(* CODESYS project Syn_Visu_3.2.0.library
   Version: 3.2.0.0
   Title: SynVisu
   Placeholder: SynVisu
   Company: Syntegon Group
   DefaultNamespace: SynVisu

Project tree, tasks and I/O mapping:
  libraries: Tc2_System, * (Beckhoff Automation GmbH)
  DUTs/
    data type E_VisuComponentType
    data type E_VisuProductState
    data type E_VisuZoneKind
    data type ST_VisuCartesian
    data type ST_VisuCartesianConfig
    data type ST_VisuCartesianState
    data type ST_VisuConveyor
    data type ST_VisuConveyorConfig
    data type ST_VisuConveyorState
    data type ST_VisuDelta
    data type ST_VisuDeltaConfig
    data type ST_VisuDeltaState
    data type ST_VisuFault
    data type ST_VisuFinger
    data type ST_VisuFingerState
    data type ST_VisuGantryMover
    data type ST_VisuLimitArea
    data type ST_VisuLoopMover
    data type ST_VisuManifest
    data type ST_VisuManifestEntry
    data type ST_VisuPlanarPose
    data type ST_VisuPose
    data type ST_VisuPosition
    data type ST_VisuProduct
    data type ST_VisuProductType
    data type ST_VisuWorkingArea
    data type ST_VisuXtsGantry
    data type ST_VisuXtsGantryConfig
    data type ST_VisuXtsGantryState
    data type ST_VisuXtsLoop
    data type ST_VisuXtsLoopConfig
    data type ST_VisuXtsLoopState
    data type ST_VisuZone
  GVLs/
    global variables VISU_GlobalConst
    global variables VISU_GlobalConst_Param
  POUs/
    function block _FB_VisuCartesian [ST]: m_ApplyConfig, m_ClearFingers, m_ClearZones, m_ComponentType, m_Configure, m_SetAxes, m_SetFault, m_SetFinger, m_SetFingerState, m_SetZone
    function block _FB_VisuComponent [ST]: m_ComponentType, m_DcTime, m_Id, m_NotifyConfigChanged, m_Register
    function block _FB_VisuConveyor [ST]: m_ApplyConfig, m_BeltPosition, m_ComponentType, m_Configure, m_FindProduct, m_GetProduct, m_LatchProduct, m_MoveProduct, m_ProductCount, m_ProductPose, m_RemoveProduct, m_RemoveProductsBeyond, m_SetBeltPosition, m_SetFault, m_SetModuloBeltPosition, m_SetProductState, m_SetProductType
    function block _FB_VisuDelta [ST]: m_ApplyConfig, m_BasePose, m_ClearFingers, m_ClearLimitArea, m_ClearZones, m_ComponentType, m_Configure, m_SetFault, m_SetFinger, m_SetFingerState, m_SetLimitArea, m_SetTcp, m_SetWorkingArea, m_SetZone
    function block _FB_VisuXtsGantry [ST]: m_ApplyConfig, m_ClearFingers, m_ClearZones, m_ComponentType, m_Configure, m_SetFault, m_SetFinger, m_SetMover, m_SetMoverCount, m_SetZone, m_SetZPosition
    function block _FB_VisuXtsLoop [ST]: m_ApplyConfig, m_ClearFingers, m_ClearZones, m_ComponentType, m_Configure, m_Perimeter, m_SetFault, m_SetFinger, m_SetMover, m_SetMoverCount, m_SetZone
    function _FC_GetVersionSynVisu [ST]
*)

// DUTs/E_VisuComponentType
{attribute 'qualified_only'}
{attribute 'strict'}
TYPE E_VisuComponentType :
(
	(* Values are part of the gateway contract: append, never renumber. *)
	NONE := 0,
	CONVEYOR := 1,
	DELTA := 2,
	XTS_GANTRY := 3,
	XTS_LOOP := 4,
	CARTESIAN := 5
) UINT;
END_TYPE

// DUTs/E_VisuProductState
{attribute 'qualified_only'}
{attribute 'strict'}
TYPE E_VisuProductState :
(
	(* Values are part of the gateway contract: append, never renumber. *)
	DETECTED := 0,
	ASSIGNED := 1,
	PICKED := 2,
	REJECTED := 3,
	PLACED := 4
) UINT;
END_TYPE

// DUTs/E_VisuZoneKind
{attribute 'qualified_only'}
{attribute 'strict'}
TYPE E_VisuZoneKind :
(
	(* Values are part of the gateway contract: append, never renumber. *)
	PICK := 1,
	PLACE := 2
) UINT;
END_TYPE

// DUTs/ST_VisuCartesian
TYPE ST_VisuCartesian :
STRUCT
	(* One visualised Cartesian robot. Register the instance's symbol path in the manifest with
	   eType := E_VisuComponentType.CARTESIAN. *)
	stConfig : ST_VisuCartesianConfig; // read at discovery and after nConfigVersion changes
	stState : ST_VisuCartesianState; // read every gateway cycle
END_STRUCT
END_TYPE

// DUTs/ST_VisuCartesianConfig
TYPE ST_VisuCartesianConfig :
STRUCT
	(* Cartesian robot: two fixed rails along local +Y, a bridge travelling in Y, a carriage on it travelling in X
	   and a vertical column (Z) ending at the gripper flange. Local frame: origin at axis X = Y = 0, Z up; the
	   flange is at (X, Y, Z). *)
	stPose : ST_VisuPose; // MCS
	fXMin : LREAL; // mm, X stroke
	fXMax : LREAL; // mm
	fYMin : LREAL; // mm, Y stroke
	fYMax : LREAL; // mm
	fZMin : LREAL; // mm, Z stroke
	fZMax : LREAL; // mm
	fRailHeight : LREAL; // mm, top of the rails above the local origin; the bridge sits on them
	nZoneCount : UINT;
	aZones : ARRAY[0..VISU_GlobalConst_Param.VISU_un_MAX_ZONES - 1] OF ST_VisuZone; // pick and place zones
	nFingerCount : UINT; // 0 = no gripper definition
	aFingers : ARRAY[0..VISU_GlobalConst_Param.VISU_un_MAX_FINGERS - 1] OF ST_VisuFinger;
END_STRUCT
END_TYPE

// DUTs/ST_VisuCartesianState
TYPE ST_VisuCartesianState :
STRUCT
	nTimestamp : ULINT; // DC time of the writing cycle, ns since 2000-01-01 (set by _FB_VisuCartesian)
	fX : LREAL; // mm, actual value: the gripper flange
	fY : LREAL; // mm, actual value
	fZ : LREAL; // mm, actual value
	bGripperActive : BOOL; // used only when no fingers are configured
	aFingerStates : ARRAY[0..VISU_GlobalConst_Param.VISU_un_MAX_FINGERS - 1] OF ST_VisuFingerState; // one per configured finger
	stFault : ST_VisuFault; // fault of the robot (set by _FB_VisuCartesian.m_SetFault)
END_STRUCT
END_TYPE

// DUTs/ST_VisuConveyor
TYPE ST_VisuConveyor :
STRUCT
	(* One visualised conveyor. Register the instance's symbol path in the manifest with
	   eType := E_VisuComponentType.CONVEYOR. *)
	stConfig : ST_VisuConveyorConfig; // read at discovery and after nConfigVersion changes
	stState : ST_VisuConveyorState; // read every gateway cycle
END_STRUCT
END_TYPE

// DUTs/ST_VisuConveyorConfig
TYPE ST_VisuConveyorConfig :
STRUCT
	stPose : ST_VisuPose; // belt start on the belt surface; local +X = conveying direction
	fLength : LREAL; // mm
	fWidth : LREAL; // mm
	nProductTypeCount : UINT;
	aProductTypes : ARRAY[0..VISU_GlobalConst_Param.VISU_un_MAX_PRODUCT_TYPES - 1] OF ST_VisuProductType;
END_STRUCT
END_TYPE

// DUTs/ST_VisuConveyorState
TYPE ST_VisuConveyorState :
STRUCT
	nTimestamp : ULINT; // DC time of the writing cycle, ns since 2000-01-01 (set by _FB_VisuConveyor)
	fBeltPosition : LREAL; // continuous belt surface position, mm, no modulo (see _FB_VisuConveyor.m_SetModuloBeltPosition)
	nProductCount : UINT; // entries [0..nProductCount-1] are evaluated
	aProducts : ARRAY[0..VISU_GlobalConst_Param.VISU_un_MAX_PRODUCTS - 1] OF ST_VisuProduct;
	stFault : ST_VisuFault; // fault of the conveyor (set by _FB_VisuConveyor.m_SetFault)
END_STRUCT
END_TYPE

// DUTs/ST_VisuDelta
TYPE ST_VisuDelta :
STRUCT
	(* One visualised Delta robot. Register the instance's symbol path in the manifest with
	   eType := E_VisuComponentType.DELTA. *)
	stConfig : ST_VisuDeltaConfig; // read at discovery and after nConfigVersion changes
	stState : ST_VisuDeltaState; // read every gateway cycle
END_STRUCT
END_TYPE

// DUTs/ST_VisuDeltaConfig
TYPE ST_VisuDeltaConfig :
STRUCT
	(* Geometry the visualisation uses to derive the arm posture from the TCP.
	   Arm 1 lies along the base's local +X; arms 2 and 3 follow counter-clockwise
	   (seen from above) at 120 deg each. *)
	stPose : ST_VisuPose; // base centre in the MCS
	fBaseRadius : LREAL; // mm, base centre to shoulder joint
	fEffectorRadius : LREAL; // mm, effector centre to lower-arm joint
	fUpperArmLength : LREAL; // mm
	fLowerArmLength : LREAL; // mm
	stWorkingArea : ST_VisuWorkingArea;
	stLimitArea : ST_VisuLimitArea; // optional box that further restricts the working area
	nZoneCount : UINT;
	aZones : ARRAY[0..VISU_GlobalConst_Param.VISU_un_MAX_ZONES - 1] OF ST_VisuZone; // pick and place zones
	nFingerCount : UINT; // 0 = no gripper definition
	aFingers : ARRAY[0..VISU_GlobalConst_Param.VISU_un_MAX_FINGERS - 1] OF ST_VisuFinger;
END_STRUCT
END_TYPE

// DUTs/ST_VisuDeltaState
TYPE ST_VisuDeltaState :
STRUCT
	nTimestamp : ULINT; // DC time of the writing cycle, ns since 2000-01-01 (set by _FB_VisuDelta.m_SetTcp)
	stActualTcp : ST_VisuPosition; // MCS, effector centre (the gripper flange); the visualisation derives the arms from it
	stSetpointTcp : ST_VisuPosition; // MCS
	aFingerStates : ARRAY[0..VISU_GlobalConst_Param.VISU_un_MAX_FINGERS - 1] OF ST_VisuFingerState; // one per configured finger
	stFault : ST_VisuFault; // fault of the robot (set by _FB_VisuDelta.m_SetFault)
END_STRUCT
END_TYPE

// DUTs/ST_VisuFault
(* Fault of a component or an XTS mover: drawn red with sMessage while bActive (contract, protocol 8). *)
TYPE ST_VisuFault :
STRUCT
	bActive : BOOL; // TRUE while the fault is active
	sMessage : STRING(80); // shown to the operator; empty shows 'Fault'
END_STRUCT
END_TYPE

// DUTs/ST_VisuFinger
TYPE ST_VisuFinger :
STRUCT
	(* One gripper finger, always drawn as a cylinder. Its frame's origin is the centre of its top face; it extends
	   along its local -Z. The grip point, where a carried product's top touches, is the centre of its bottom face. *)
	fDiameter : LREAL; // mm
	fHeight : LREAL; // mm
END_STRUCT
END_TYPE

// DUTs/ST_VisuFingerState
TYPE ST_VisuFingerState :
STRUCT
	stPose : ST_VisuPose; // MCS, absolute: pose of the finger's frame (centre of its top face)
	bActive : BOOL; // the finger grips
END_STRUCT
END_TYPE

// DUTs/ST_VisuGantryMover
TYPE ST_VisuGantryMover :
STRUCT
	nId : UDINT; // unique within the gantry, > 0; referenced by a carried product's nMoverId
	bValid : BOOL; // invalid entries are not shown
	fPosition : LREAL; // mm along the track (local +Y), actual value
	fX : LREAL; // mm, X axis on the mover, actual value
	bGripperActive : BOOL; // used only when no fingers are configured
	aFingerStates : ARRAY[0..VISU_GlobalConst_Param.VISU_un_MAX_FINGERS - 1] OF ST_VisuFingerState; // one per configured finger
	stFault : ST_VisuFault; // fault of this mover
END_STRUCT
END_TYPE

// DUTs/ST_VisuLimitArea
TYPE ST_VisuLimitArea :
STRUCT
	(* Axis-aligned box in the robot frame (relative to the base centre, turned with the robot's pose) that further
	   restricts the working area, e.g. so that neighbouring robots cannot collide. *)
	fXMin : LREAL; // mm
	fXMax : LREAL; // mm
	fYMin : LREAL; // mm
	fYMax : LREAL; // mm
	fZMin : LREAL; // mm relative to the base (below the base: negative)
	fZMax : LREAL; // mm relative to the base
	bActive : BOOL; // FALSE: no limit area, the box is not drawn
END_STRUCT
END_TYPE

// DUTs/ST_VisuLoopMover
TYPE ST_VisuLoopMover :
STRUCT
	nId : UDINT; // unique within the loop, > 0; referenced by a carried product's nMoverId
	bValid : BOOL; // invalid entries are not shown
	fPosition : LREAL; // mm along the loop from the start of the lower straight, in the conveying direction
	aFingerStates : ARRAY[0..VISU_GlobalConst_Param.VISU_un_MAX_FINGERS - 1] OF ST_VisuFingerState; // one per configured finger
	stFault : ST_VisuFault; // fault of this mover
END_STRUCT
END_TYPE

// DUTs/ST_VisuManifest
TYPE ST_VisuManifest :
STRUCT
	(* Discovery entry point. The application declares one instance at the fixed symbol
	   GVL_Visu.stManifest; the gateway starts reading there. *)
	nProtocolVersion : UINT := VISU_GlobalConst.VISU_un_PROTOCOL_VERSION;
	(* Increment after any change to the manifest or to a component's stConfig. *)
	nConfigVersion : UDINT := 1;
	nCount : UINT; // entries [0..nCount-1] are evaluated
	aEntries : ARRAY[0..VISU_GlobalConst_Param.VISU_un_MAX_MANIFEST_ENTRIES - 1] OF ST_VisuManifestEntry;
END_STRUCT
END_TYPE

// DUTs/ST_VisuManifestEntry
TYPE ST_VisuManifestEntry :
STRUCT
	nId : UDINT; // unique within the manifest, > 0; used for all cross-references
	eType : E_VisuComponentType;
	sName : STRING(80); // display name
	sPath : STRING(255); // symbol path of the ST_VisuConveyor / ST_VisuDelta instance, e.g. 'MAIN.stInfeed'
END_STRUCT
END_TYPE

// DUTs/ST_VisuPlanarPose
TYPE ST_VisuPlanarPose :
STRUCT
	(* Position plus rotation about Z in the MCS, used for TCPs and product latch poses. *)
	fX : LREAL; // mm
	fY : LREAL; // mm
	fZ : LREAL; // mm
	fRz : LREAL; // degrees
END_STRUCT
END_TYPE

// DUTs/ST_VisuPose
TYPE ST_VisuPose :
STRUCT
	(* Pose in the MCS: right-handed, Z up, X in product flow direction.
	   Rotation order R = Rz(fRz) * Ry(fRy) * Rx(fRx). *)
	fX : LREAL; // mm
	fY : LREAL; // mm
	fZ : LREAL; // mm
	fRx : LREAL; // degrees
	fRy : LREAL; // degrees
	fRz : LREAL; // degrees
END_STRUCT
END_TYPE

// DUTs/ST_VisuPosition
TYPE ST_VisuPosition :
STRUCT
	(* A point in the MCS, e.g. a Delta's TCP. *)
	fX : LREAL; // mm
	fY : LREAL; // mm
	fZ : LREAL; // mm
END_STRUCT
END_TYPE

// DUTs/ST_VisuProduct
TYPE ST_VisuProduct :
STRUCT
	nId : UDINT;
	bValid : BOOL; // invalid entries are not shown
	stLatchPose : ST_VisuPlanarPose; // MCS, bottom centre of the product at latch time
	fLatchBeltPosition : LREAL; // conveyor fBeltPosition at latch time, mm
	eState : E_VisuProductState;
	nRobotId : UDINT; // manifest id of the assigned robot, 0 = none
	nMoverId : UDINT; // mover of an XTS gantry or loop carrying the product, 0 = none
	nFingerId : UDINT; // gripper finger (1-based) the product hangs from while picked, 0 = the gripper flange
	nProductType : UDINT; // id in the conveyor's aProductTypes
END_STRUCT
END_TYPE

// DUTs/ST_VisuProductType
TYPE ST_VisuProductType :
STRUCT
	nId : UDINT;
	fLength : LREAL; // mm, along the conveying direction
	fWidth : LREAL; // mm
	fHeight : LREAL; // mm
END_STRUCT
END_TYPE

// DUTs/ST_VisuWorkingArea
TYPE ST_VisuWorkingArea :
STRUCT
	(* Limit shape the PLC enforces: vertical cylinder in the robot frame, optional cone below. *)
	fRadius : LREAL; // mm
	fZMin : LREAL; // mm relative to the base (below the base: negative)
	fZMax : LREAL; // mm relative to the base
	fConeHeight : LREAL; // mm below fZMin; 0 = no cone
	fConeBottomRadius : LREAL; // mm
END_STRUCT
END_TYPE

// DUTs/ST_VisuXtsGantry
TYPE ST_VisuXtsGantry :
STRUCT
	(* One visualised XTS gantry (e.g. IDH). Register the instance's symbol path in the manifest with
	   eType := E_VisuComponentType.XTS_GANTRY. *)
	stConfig : ST_VisuXtsGantryConfig; // read at discovery and after nConfigVersion changes
	stState : ST_VisuXtsGantryState; // read every gateway cycle
END_STRUCT
END_TYPE

// DUTs/ST_VisuXtsGantryConfig
TYPE ST_VisuXtsGantryConfig :
STRUCT
	(* Straight XTS track of equal modules, carried by a common Z axis; every mover carries an X axis with a
	   gripper flange at its end. Local frame: origin at the track start on top of the movers with Z = 0; the track runs
	   along local +Y, the X axes along local +X, the Z axis along local +Z (up). *)
	stPose : ST_VisuPose; // MCS
	nModuleCount : UINT; // track modules in a row
	fModuleLength : LREAL; // mm, length of one module
	fXMin : LREAL; // mm, X stroke
	fXMax : LREAL; // mm
	fZMin : LREAL; // mm, Z stroke
	fZMax : LREAL; // mm
	fToolOffsetX : LREAL; // mm, gripper flange ahead of the X axis zero along local +X
	fToolOffsetZ : LREAL; // mm, gripper flange relative to the mover top (below: negative)
	fMoverLength : LREAL; // mm, along the track
	fMoverWidth : LREAL; // mm
	nZoneCount : UINT;
	aZones : ARRAY[0..VISU_GlobalConst_Param.VISU_un_MAX_ZONES - 1] OF ST_VisuZone; // pick and place zones
	nFingerCount : UINT; // fingers of every mover's gripper, 0 = no gripper definition
	aFingers : ARRAY[0..VISU_GlobalConst_Param.VISU_un_MAX_FINGERS - 1] OF ST_VisuFinger;
END_STRUCT
END_TYPE

// DUTs/ST_VisuXtsGantryState
TYPE ST_VisuXtsGantryState :
STRUCT
	nTimestamp : ULINT; // DC time of the writing cycle, ns since 2000-01-01 (set by _FB_VisuXtsGantry)
	fZ : LREAL; // mm, common Z axis, actual value
	nMoverCount : UINT; // entries [0..nMoverCount-1] are evaluated
	aMovers : ARRAY[0..VISU_GlobalConst_Param.VISU_un_MAX_MOVERS - 1] OF ST_VisuGantryMover;
	stFault : ST_VisuFault; // fault of the whole gantry (set by _FB_VisuXtsGantry.m_SetFault)
END_STRUCT
END_TYPE

// DUTs/ST_VisuXtsLoop
TYPE ST_VisuXtsLoop :
STRUCT
	(* One visualised XTS loop (e.g. Fxx). Register the instance's symbol path in the manifest with
	   eType := E_VisuComponentType.XTS_LOOP. *)
	stConfig : ST_VisuXtsLoopConfig; // read at discovery and after nConfigVersion changes
	stState : ST_VisuXtsLoopState; // read every gateway cycle
END_STRUCT
END_TYPE

// DUTs/ST_VisuXtsLoopConfig
TYPE ST_VisuXtsLoopConfig :
STRUCT
	(* Closed XTS loop: two straights joined by two 180 deg curves (drawn as semicircles), standing in the local X-Z
	   plane. Local frame: origin at the start of the lower straight, which runs along local +X in the conveying
	   direction; the upper straight lies at +2 * fCurveRadius in Z. *)
	stPose : ST_VisuPose; // MCS
	fStraightLength : LREAL; // mm
	fCurveRadius : LREAL; // mm
	fToolOffset : LREAL; // mm, gripper flange (tool point) of a mover outwards from the track
	fMoverLength : LREAL; // mm, along the track
	fMoverWidth : LREAL; // mm
	nZoneCount : UINT;
	aZones : ARRAY[0..VISU_GlobalConst_Param.VISU_un_MAX_ZONES - 1] OF ST_VisuZone; // pick and place zones
	nFingerCount : UINT; // fingers of every mover's gripper, 0 = no gripper definition
	aFingers : ARRAY[0..VISU_GlobalConst_Param.VISU_un_MAX_FINGERS - 1] OF ST_VisuFinger;
END_STRUCT
END_TYPE

// DUTs/ST_VisuXtsLoopState
TYPE ST_VisuXtsLoopState :
STRUCT
	nTimestamp : ULINT; // DC time of the writing cycle, ns since 2000-01-01 (set by _FB_VisuXtsLoop)
	nMoverCount : UINT; // entries [0..nMoverCount-1] are evaluated
	aMovers : ARRAY[0..VISU_GlobalConst_Param.VISU_un_MAX_MOVERS - 1] OF ST_VisuLoopMover;
	stFault : ST_VisuFault; // fault of the whole loop (set by _FB_VisuXtsLoop.m_SetFault)
END_STRUCT
END_TYPE

// DUTs/ST_VisuZone
TYPE ST_VisuZone :
STRUCT
	nConveyorId : UDINT; // manifest id of the conveyor
	fStart : LREAL; // mm along the conveyor's local X (belt coordinates, not MCS)
	fEnd : LREAL; // mm along the conveyor's local X
	eKind : E_VisuZoneKind;
	(* mm before fEnd, against the conveying direction: the robot may allocate products in the zone only up to
	   fEnd - fAllocationOffset, so it does not move out of the zone while approaching. 0 = no allocation limit. *)
	fAllocationOffset : LREAL;
END_STRUCT
END_TYPE

// GVLs/VISU_GlobalConst
(****************************************************************************************************<br>
© Syntegon Group.<br>
All rights reserved, also regarding any disposal, exploitation, reproduction, editing, distribution,<br>
as well as in the event of applications for industrial property rights.<br>
*****************************************************************************************************<br>
DESCRIPTION:<br>
Global constants of the Syn_Visu library.<br>
****************************************************************************************************)
{attribute 'qualified_only'}
VAR_GLOBAL CONSTANT
	(* Version of the PLC <-> gateway contract. The gateway refuses to read a PLC whose manifest
	   reports a different value. Bump together with PROTOCOL_VERSION in the gateway.
	   2: the Delta reports only its TCP; the visualisation derives the arm posture.
	   3: work area renamed to working area, windows to zones.
	   4: XTS gantry and XTS loop, product nMoverId, fEncoder renamed to fBeltPosition.
	   5: Cartesian robot.
	   6: Delta limit area, zone allocation offset.
	   7: gripper fingers; tool rotations (Delta rz, IDH C, Cartesian C/A and tool length) removed.
	   8: faults of components and XTS movers (stFault). *)
	VISU_un_PROTOCOL_VERSION			: UINT := 8;
	VISU_lr_DEG_TO_RAD					: LREAL := 0.017453292519943295;	// [rad/deg] pi / 180
END_VAR

// GVLs/VISU_GlobalConst_Param
(****************************************************************************************************<br>
© Syntegon Group.<br>
All rights reserved, also regarding any disposal, exploitation, reproduction, editing, distribution,<br>
as well as in the event of applications for industrial property rights.<br>
*****************************************************************************************************<br>
DESCRIPTION:<br>
Library parameters of Syn_Visu: array sizes of the interface structures.<br>
****************************************************************************************************)
{attribute 'qualified_only'}
VAR_GLOBAL CONSTANT
	VISU_un_MAX_MANIFEST_ENTRIES		: UINT := 32;	// [-] components in the manifest
	VISU_un_MAX_PRODUCTS				: UINT := 128;	// [-] products per conveyor
	VISU_un_MAX_PRODUCT_TYPES			: UINT := 8;	// [-] product types per conveyor
	VISU_un_MAX_ZONES					: UINT := 8;	// [-] zones per robot
	VISU_un_MAX_MOVERS					: UINT := 40;	// [-] movers per XTS gantry or loop
	VISU_un_MAX_FINGERS					: UINT := 8;	// [-] fingers per gripper
END_VAR

// POUs/_FB_VisuCartesian
(****************************************************************************************************<br>
© Syntegon Group.<br>
All rights reserved, also regarding any disposal, exploitation, reproduction, editing, distribution,<br>
as well as in the event of applications for industrial property rights.<br>
*****************************************************************************************************<br>
DESCRIPTION:<br>
One visualised Cartesian robot: linear X, Y, Z axes ending at a gripper flange. Typical cycle:<br>
  fb_Cartesian.m_Register(vio_Manifest := GVL_Visu.stManifest, vi_udn_Id := 40, vi_str_Name := 'Cartesian',<br>
      vi_str_Path := 'MAIN.fb_Cartesian.vo_Visu');<br>
  fb_Cartesian.m_Configure(vi_Pose := RobotPose, vi_lr_XMin := 0, vi_lr_XMax := 1200, vi_lr_YMin := 0,<br>
      vi_lr_YMax := 1000, vi_lr_ZMin := -600, vi_lr_ZMax := 0, vi_lr_RailHeight := 1200);<br>
  fb_Cartesian.m_SetFinger(vi_un_Finger := 1, vi_lr_Diameter := 40, vi_lr_Height := 40);<br>
  fb_Cartesian.m_SetZone(vi_udn_ConveyorId := 7, vi_e_Kind := E_VisuZoneKind.PICK, vi_lr_Start := 1000, vi_lr_End := 2000);<br>
  fb_Cartesian.m_SetAxes(vi_lr_X := ..., vi_lr_Y := ..., vi_lr_Z := ...);<br>
  fb_Cartesian.m_SetFingerState(vi_un_Finger := 1, vi_Pose := CupPose, vi_b_Active := b_Vacuum);<br>
Only actual values are reported; tool rotations (e.g. C and A) show only through the finger poses, absolute in<br>
the MCS. The config methods may be called every cycle; the config version only changes when a value does.<br>
*****************************************************************************************************<br>
OUTPUT VALUES:<br>
vo_Visu is the contract structure the gateway reads at the path given to m_Register. Do not write it.<br>
*****************************************************************************************************<br>
VERSION         ¦ DATE       ¦ NAME      ¦ CHANGE<br>
Syn_Visu 3.0.0  ¦ 2026-10-31 ¦ J.Willner ¦ Naming and layout after the TCAT programming guideline<br>
****************************************************************************************************)
FUNCTION_BLOCK _FB_VisuCartesian EXTENDS _FB_VisuComponent
VAR_OUTPUT
	vo_Visu								: ST_VisuCartesian;	// contract structure read by the gateway
END_VAR

(****************************************************************************************************<br>
© Syntegon Group.<br>
All rights reserved, also regarding any disposal, exploitation, reproduction, editing, distribution,<br>
as well as in the event of applications for industrial property rights.<br>
*****************************************************************************************************<br>
DESCRIPTION:<br>
Takes over vio_New and increments the config version if it differs from the current config. TRUE if changed.<br>
****************************************************************************************************)
METHOD PRIVATE m_ApplyConfig : BOOL
VAR_IN_OUT
	vio_New								: ST_VisuCartesianConfig;
END_VAR
m_ApplyConfig := Tc2_System.MEMCMP(ADR(vio_New), ADR(vo_Visu.stConfig), SIZEOF(vio_New)) <> 0;
IF m_ApplyConfig THEN
	vo_Visu.stConfig := vio_New;
	m_NotifyConfigChanged();
END_IF
END_METHOD

(****************************************************************************************************<br>
© Syntegon Group.<br>
All rights reserved, also regarding any disposal, exploitation, reproduction, editing, distribution,<br>
as well as in the event of applications for industrial property rights.<br>
*****************************************************************************************************<br>
DESCRIPTION:<br>
Removes the gripper definition. TRUE if there was one.<br>
****************************************************************************************************)
METHOD m_ClearFingers : BOOL
VAR
	TempNew								: ST_VisuCartesianConfig;
	TempEmpty							: ST_VisuFinger;
	un_TempIndex						: UINT;
END_VAR
TempNew := vo_Visu.stConfig;
FOR un_TempIndex := 0 TO VISU_GlobalConst_Param.VISU_un_MAX_FINGERS - 1 DO
	TempNew.aFingers[un_TempIndex] := TempEmpty;
END_FOR
TempNew.nFingerCount := 0;
m_ClearFingers := m_ApplyConfig(TempNew);
END_METHOD

(****************************************************************************************************<br>
© Syntegon Group.<br>
All rights reserved, also regarding any disposal, exploitation, reproduction, editing, distribution,<br>
as well as in the event of applications for industrial property rights.<br>
*****************************************************************************************************<br>
DESCRIPTION:<br>
Removes all pick and place zones. TRUE if there were any.<br>
****************************************************************************************************)
METHOD m_ClearZones : BOOL
VAR
	TempNew								: ST_VisuCartesianConfig;
	TempEmpty							: ST_VisuZone;
	un_TempIndex						: UINT;
END_VAR
TempNew := vo_Visu.stConfig;
FOR un_TempIndex := 0 TO VISU_GlobalConst_Param.VISU_un_MAX_ZONES - 1 DO
	TempNew.aZones[un_TempIndex] := TempEmpty;
END_FOR
TempNew.nZoneCount := 0;
m_ClearZones := m_ApplyConfig(TempNew);
END_METHOD

(****************************************************************************************************<br>
© Syntegon Group.<br>
All rights reserved, also regarding any disposal, exploitation, reproduction, editing, distribution,<br>
as well as in the event of applications for industrial property rights.<br>
*****************************************************************************************************<br>
DESCRIPTION:<br>
Manifest type: Cartesian robot.<br>
****************************************************************************************************)
METHOD PROTECTED m_ComponentType : E_VisuComponentType
m_ComponentType := E_VisuComponentType.CARTESIAN;
END_METHOD

(****************************************************************************************************<br>
© Syntegon Group.<br>
All rights reserved, also regarding any disposal, exploitation, reproduction, editing, distribution,<br>
as well as in the event of applications for industrial property rights.<br>
*****************************************************************************************************<br>
DESCRIPTION:<br>
Sets pose, strokes and rail height. TRUE if anything changed.<br>
****************************************************************************************************)
METHOD m_Configure : BOOL
VAR_INPUT
	vi_Pose								: ST_VisuPose;	// MCS, axis origin X = Y = 0 with Z up
	vi_lr_XMin							: LREAL;	// [mm]
	vi_lr_XMax							: LREAL;	// [mm]
	vi_lr_YMin							: LREAL;	// [mm]
	vi_lr_YMax							: LREAL;	// [mm]
	vi_lr_ZMin							: LREAL;	// [mm]
	vi_lr_ZMax							: LREAL;	// [mm]
	vi_lr_RailHeight					: LREAL;	// [mm] top of the rails above the local origin
END_VAR
VAR
	TempNew								: ST_VisuCartesianConfig;
END_VAR
TempNew := vo_Visu.stConfig;
TempNew.stPose := vi_Pose;
TempNew.fXMin := vi_lr_XMin;
TempNew.fXMax := vi_lr_XMax;
TempNew.fYMin := vi_lr_YMin;
TempNew.fYMax := vi_lr_YMax;
TempNew.fZMin := vi_lr_ZMin;
TempNew.fZMax := vi_lr_ZMax;
TempNew.fRailHeight := vi_lr_RailHeight;
m_Configure := m_ApplyConfig(TempNew);
END_METHOD

(****************************************************************************************************<br>
© Syntegon Group.<br>
All rights reserved, also regarding any disposal, exploitation, reproduction, editing, distribution,<br>
as well as in the event of applications for industrial property rights.<br>
*****************************************************************************************************<br>
DESCRIPTION:<br>
Reports the axes' actual values and the gripper. Call once per cycle; it also stamps the state with the<br>
cycle's DC time.<br>
****************************************************************************************************)
METHOD m_SetAxes : BOOL
VAR_INPUT
	vi_lr_X								: LREAL;	// [mm]
	vi_lr_Y								: LREAL;	// [mm]
	vi_lr_Z								: LREAL;	// [mm]
	vi_b_GripperActive					: BOOL := FALSE;	// used only when no fingers are configured
END_VAR
vo_Visu.stState.fX := vi_lr_X;
vo_Visu.stState.fY := vi_lr_Y;
vo_Visu.stState.fZ := vi_lr_Z;
vo_Visu.stState.bGripperActive := vi_b_GripperActive;
vo_Visu.stState.nTimestamp := m_DcTime();
m_SetAxes := TRUE;
END_METHOD

(****************************************************************************************************<br>
© Syntegon Group.<br>
All rights reserved, also regarding any disposal, exploitation, reproduction, editing, distribution,<br>
as well as in the event of applications for industrial property rights.<br>
*****************************************************************************************************<br>
DESCRIPTION:<br>
Sets or clears the fault of the robot: drawn red with the message while active. The fault stays until it<br>
is cleared with m_SetFault(vi_b_Active := FALSE, vi_str_Message := ''). TRUE.<br>
****************************************************************************************************)
METHOD m_SetFault : BOOL
VAR_INPUT
	vi_b_Active							: BOOL;	// TRUE: fault active
	vi_str_Message						: STRING(80);	// shown to the operator; empty shows 'Fault'
END_VAR
vo_Visu.stState.stFault.bActive := vi_b_Active;
vo_Visu.stState.stFault.sMessage := vi_str_Message;
m_SetFault := TRUE;
END_METHOD

(****************************************************************************************************<br>
© Syntegon Group.<br>
All rights reserved, also regarding any disposal, exploitation, reproduction, editing, distribution,<br>
as well as in the event of applications for industrial property rights.<br>
*****************************************************************************************************<br>
DESCRIPTION:<br>
Defines gripper finger vi_un_Finger (1-based): a cylinder hanging from the finger's pose along its local -Z.<br>
The finger count grows to vi_un_Finger.<br>
*****************************************************************************************************<br>
OUTPUT VALUES:<br>
FALSE outside 1..VISU_GlobalConst_Param.VISU_un_MAX_FINGERS.<br>
****************************************************************************************************)
METHOD m_SetFinger : BOOL
VAR_INPUT
	vi_un_Finger						: UINT;	// [-] 1-based, as a product's nFingerId
	vi_lr_Diameter						: LREAL;	// [mm]
	vi_lr_Height						: LREAL;	// [mm] along the finger's local -Z
END_VAR
VAR
	TempNew								: ST_VisuCartesianConfig;
END_VAR
m_SetFinger := FALSE;
IF vi_un_Finger = 0 OR vi_un_Finger > VISU_GlobalConst_Param.VISU_un_MAX_FINGERS THEN
	RETURN;
END_IF
TempNew := vo_Visu.stConfig;
TempNew.aFingers[vi_un_Finger - 1].fDiameter := vi_lr_Diameter;
TempNew.aFingers[vi_un_Finger - 1].fHeight := vi_lr_Height;
TempNew.nFingerCount := MAX(TempNew.nFingerCount, vi_un_Finger);
m_ApplyConfig(TempNew);
m_SetFinger := TRUE;
END_METHOD

(****************************************************************************************************<br>
© Syntegon Group.<br>
All rights reserved, also regarding any disposal, exploitation, reproduction, editing, distribution,<br>
as well as in the event of applications for industrial property rights.<br>
*****************************************************************************************************<br>
DESCRIPTION:<br>
Reports finger vi_un_Finger (1-based): the pose of its frame (centre of its top face), absolute in the MCS,<br>
and whether it grips. Call once per cycle per configured finger.<br>
*****************************************************************************************************<br>
OUTPUT VALUES:<br>
FALSE outside 1..VISU_GlobalConst_Param.VISU_un_MAX_FINGERS.<br>
****************************************************************************************************)
METHOD m_SetFingerState : BOOL
VAR_INPUT
	vi_un_Finger						: UINT;	// [-] 1-based
	vi_Pose								: ST_VisuPose;	// MCS
	vi_b_Active							: BOOL;	// TRUE while the finger grips
END_VAR
m_SetFingerState := vi_un_Finger > 0 AND vi_un_Finger <= VISU_GlobalConst_Param.VISU_un_MAX_FINGERS;
IF m_SetFingerState THEN
	vo_Visu.stState.aFingerStates[vi_un_Finger - 1].stPose := vi_Pose;
	vo_Visu.stState.aFingerStates[vi_un_Finger - 1].bActive := vi_b_Active;
END_IF
END_METHOD

(****************************************************************************************************<br>
© Syntegon Group.<br>
All rights reserved, also regarding any disposal, exploitation, reproduction, editing, distribution,<br>
as well as in the event of applications for industrial property rights.<br>
*****************************************************************************************************<br>
DESCRIPTION:<br>
Adds a pick or place zone, or updates the one for the same conveyor and kind.<br>
*****************************************************************************************************<br>
OUTPUT VALUES:<br>
FALSE for vi_udn_ConveyorId = 0 or a full list.<br>
****************************************************************************************************)
METHOD m_SetZone : BOOL
VAR_INPUT
	vi_udn_ConveyorId					: UDINT;	// [-] manifest id of the conveyor
	vi_e_Kind							: E_VisuZoneKind;
	vi_lr_Start							: LREAL;	// [mm] along the conveyor from its start (belt coordinates, not MCS)
	vi_lr_End							: LREAL;	// [mm] along the conveyor from its start
	vi_lr_AllocationOffset				: LREAL := 0;	// [mm] before vi_lr_End up to which products may be allocated; 0 = no limit
END_VAR
VAR
	TempNew								: ST_VisuCartesianConfig;
	un_TempIndex						: UINT;
END_VAR
m_SetZone := FALSE;
IF vi_udn_ConveyorId = 0 THEN
	RETURN;
END_IF
TempNew := vo_Visu.stConfig;
un_TempIndex := 0;
(* ST evaluates both operands of AND: test the index before reading the array. *)
WHILE un_TempIndex < TempNew.nZoneCount DO
	IF TempNew.aZones[un_TempIndex].nConveyorId = vi_udn_ConveyorId AND TempNew.aZones[un_TempIndex].eKind = vi_e_Kind THEN
		EXIT;
	END_IF
	un_TempIndex := un_TempIndex + 1;
END_WHILE
IF un_TempIndex >= VISU_GlobalConst_Param.VISU_un_MAX_ZONES THEN
	RETURN;
END_IF
IF un_TempIndex = TempNew.nZoneCount THEN
	TempNew.nZoneCount := TempNew.nZoneCount + 1;
END_IF
TempNew.aZones[un_TempIndex].nConveyorId := vi_udn_ConveyorId;
TempNew.aZones[un_TempIndex].eKind := vi_e_Kind;
TempNew.aZones[un_TempIndex].fStart := vi_lr_Start;
TempNew.aZones[un_TempIndex].fEnd := vi_lr_End;
TempNew.aZones[un_TempIndex].fAllocationOffset := vi_lr_AllocationOffset;
m_ApplyConfig(TempNew);
m_SetZone := TRUE;
END_METHOD

END_FUNCTION_BLOCK

// POUs/_FB_VisuComponent
(****************************************************************************************************<br>
© Syntegon Group.<br>
All rights reserved, also regarding any disposal, exploitation, reproduction, editing, distribution,<br>
as well as in the event of applications for industrial property rights.<br>
*****************************************************************************************************<br>
DESCRIPTION:<br>
Base of every visualised component (_FB_VisuConveyor, _FB_VisuDelta, ...). Handles the manifest entry,<br>
the config version and the DC timestamps. Not used directly.<br>
*****************************************************************************************************<br>
VERSION         ¦ DATE       ¦ NAME      ¦ CHANGE<br>
Syn_Visu 3.0.0  ¦ 2026-10-31 ¦ J.Willner ¦ Naming and layout after the TCAT programming guideline<br>
****************************************************************************************************)
FUNCTION_BLOCK ABSTRACT _FB_VisuComponent
VAR
	RefManifest							: REFERENCE TO ST_VisuManifest;	// set by m_Register
	udn_ComponentId						: UDINT;	// [-] manifest id, 0 = not registered
END_VAR

(****************************************************************************************************<br>
© Syntegon Group.<br>
All rights reserved, also regarding any disposal, exploitation, reproduction, editing, distribution,<br>
as well as in the event of applications for industrial property rights.<br>
*****************************************************************************************************<br>
DESCRIPTION:<br>
Manifest type of the component. Overridden by every derived FB.<br>
****************************************************************************************************)
METHOD PROTECTED m_ComponentType : E_VisuComponentType
m_ComponentType := E_VisuComponentType.NONE;
END_METHOD

(****************************************************************************************************<br>
© Syntegon Group.<br>
All rights reserved, also regarding any disposal, exploitation, reproduction, editing, distribution,<br>
as well as in the event of applications for industrial property rights.<br>
*****************************************************************************************************<br>
DESCRIPTION:<br>
Distributed-clock time of the calling task's current cycle in ns since 2000-01-01; 0 if unknown.<br>
****************************************************************************************************)
METHOD PROTECTED m_DcTime : ULINT
VAR
	dn_TempTaskIndex					: DINT;
END_VAR
dn_TempTaskIndex := Tc2_System.GETCURTASKINDEXEX();
IF dn_TempTaskIndex > 0 THEN
	m_DcTime := LINT_TO_ULINT(TwinCAT_SystemInfoVarList._TaskInfo[dn_TempTaskIndex].DcTaskTime);
ELSE
	m_DcTime := 0;
END_IF
END_METHOD

(****************************************************************************************************<br>
© Syntegon Group.<br>
All rights reserved, also regarding any disposal, exploitation, reproduction, editing, distribution,<br>
as well as in the event of applications for industrial property rights.<br>
*****************************************************************************************************<br>
DESCRIPTION:<br>
Manifest id given to m_Register; 0 while not registered.<br>
****************************************************************************************************)
METHOD m_Id : UDINT
m_Id := udn_ComponentId;
END_METHOD

(****************************************************************************************************<br>
© Syntegon Group.<br>
All rights reserved, also regarding any disposal, exploitation, reproduction, editing, distribution,<br>
as well as in the event of applications for industrial property rights.<br>
*****************************************************************************************************<br>
DESCRIPTION:<br>
Increments the manifest's nConfigVersion so the gateway re-reads the config. No effect before m_Register.<br>
****************************************************************************************************)
METHOD PROTECTED m_NotifyConfigChanged : BOOL
m_NotifyConfigChanged := __ISVALIDREF(RefManifest);
IF m_NotifyConfigChanged THEN
	RefManifest.nConfigVersion := RefManifest.nConfigVersion + 1;
END_IF
END_METHOD

(****************************************************************************************************<br>
© Syntegon Group.<br>
All rights reserved, also regarding any disposal, exploitation, reproduction, editing, distribution,<br>
as well as in the event of applications for industrial property rights.<br>
*****************************************************************************************************<br>
DESCRIPTION:<br>
Adds this component to the manifest; increments nConfigVersion when the entry is new.<br>
Idempotent: call it every cycle, which also keeps the manifest reference valid after an online change.<br>
*****************************************************************************************************<br>
OUTPUT VALUES:<br>
FALSE for vi_udn_Id = 0, an id already used by a different entry, or a full manifest.<br>
****************************************************************************************************)
METHOD m_Register : BOOL
VAR_IN_OUT
	vio_Manifest						: ST_VisuManifest;	// GVL_Visu.stManifest of the application
END_VAR
VAR_INPUT
	vi_udn_Id							: UDINT;	// [-] unique, > 0
	vi_str_Name							: STRING(80);	// display name
	vi_str_Path							: STRING(255);	// symbol path of this instance's vo_Visu, e.g. 'MAIN.fb_Infeed.vo_Visu'
END_VAR
VAR
	e_TempType							: E_VisuComponentType;
	un_TempIndex						: UINT;
END_VAR
m_Register := FALSE;
RefManifest REF= vio_Manifest;
(* Always report the contract version of the library actually running, also after an online change. *)
vio_Manifest.nProtocolVersion := VISU_GlobalConst.VISU_un_PROTOCOL_VERSION;
e_TempType := m_ComponentType();
IF vi_udn_Id = 0 OR e_TempType = E_VisuComponentType.NONE THEN
	RETURN;
END_IF

(* An existing entry with the same id must match exactly. *)
un_TempIndex := 0;
WHILE un_TempIndex < vio_Manifest.nCount AND un_TempIndex < VISU_GlobalConst_Param.VISU_un_MAX_MANIFEST_ENTRIES DO
	IF vio_Manifest.aEntries[un_TempIndex].nId = vi_udn_Id THEN
		m_Register := vio_Manifest.aEntries[un_TempIndex].eType = e_TempType
					AND vio_Manifest.aEntries[un_TempIndex].sName = vi_str_Name
					AND vio_Manifest.aEntries[un_TempIndex].sPath = vi_str_Path;
		IF m_Register THEN
			udn_ComponentId := vi_udn_Id;
		END_IF
		RETURN;
	END_IF
	un_TempIndex := un_TempIndex + 1;
END_WHILE

(* New entry. *)
IF vio_Manifest.nCount >= VISU_GlobalConst_Param.VISU_un_MAX_MANIFEST_ENTRIES THEN
	RETURN;
END_IF
vio_Manifest.aEntries[vio_Manifest.nCount].nId := vi_udn_Id;
vio_Manifest.aEntries[vio_Manifest.nCount].eType := e_TempType;
vio_Manifest.aEntries[vio_Manifest.nCount].sName := vi_str_Name;
vio_Manifest.aEntries[vio_Manifest.nCount].sPath := vi_str_Path;
vio_Manifest.nCount := vio_Manifest.nCount + 1;
vio_Manifest.nConfigVersion := vio_Manifest.nConfigVersion + 1;
udn_ComponentId := vi_udn_Id;
m_Register := TRUE;
END_METHOD

END_FUNCTION_BLOCK

// POUs/_FB_VisuConveyor
(****************************************************************************************************<br>
© Syntegon Group.<br>
All rights reserved, also regarding any disposal, exploitation, reproduction, editing, distribution,<br>
as well as in the event of applications for industrial property rights.<br>
*****************************************************************************************************<br>
DESCRIPTION:<br>
One visualised conveyor. Typical cycle:<br>
  fb_Infeed.m_Register(vio_Manifest := GVL_Visu.stManifest, vi_udn_Id := 1, vi_str_Name := 'Infeed',<br>
      vi_str_Path := 'MAIN.fb_Infeed.vo_Visu');<br>
  fb_Infeed.m_Configure(vi_Pose := BeltPose, vi_lr_Length := 5000, vi_lr_Width := 400);<br>
  fb_Infeed.m_SetProductType(vi_udn_Id := 1, vi_lr_Length := 120, vi_lr_Width := 80, vi_lr_Height := 40);<br>
  fb_Infeed.m_SetBeltPosition(lr_AxisPosition);  // or m_SetModuloBeltPosition for a modulo axis<br>
  IF b_Latched THEN fb_Infeed.m_LatchProduct(vi_udn_Id := udn_NextId, vi_LatchPose := LatchPose, vi_udn_ProductType := 1); END_IF<br>
m_Configure and m_SetProductType may be called every cycle; the config version only changes when a value does.<br>
*****************************************************************************************************<br>
OUTPUT VALUES:<br>
vo_Visu is the contract structure the gateway reads at the path given to m_Register. Do not write it.<br>
*****************************************************************************************************<br>
VERSION         ¦ DATE       ¦ NAME      ¦ CHANGE<br>
Syn_Visu 3.0.0  ¦ 2026-10-31 ¦ J.Willner ¦ Naming and layout after the TCAT programming guideline<br>
****************************************************************************************************)
FUNCTION_BLOCK _FB_VisuConveyor EXTENDS _FB_VisuComponent
VAR_OUTPUT
	vo_Visu								: ST_VisuConveyor;	// contract structure read by the gateway
END_VAR
VAR
	lr_LastModuloPosition				: LREAL;	// [mm] modulo position of the previous cycle
	b_ModuloInitialised					: BOOL;
END_VAR

(****************************************************************************************************<br>
© Syntegon Group.<br>
All rights reserved, also regarding any disposal, exploitation, reproduction, editing, distribution,<br>
as well as in the event of applications for industrial property rights.<br>
*****************************************************************************************************<br>
DESCRIPTION:<br>
Takes over vio_New and increments the config version if it differs from the current config. TRUE if changed.<br>
****************************************************************************************************)
METHOD PRIVATE m_ApplyConfig : BOOL
VAR_IN_OUT
	vio_New								: ST_VisuConveyorConfig;
END_VAR
m_ApplyConfig := Tc2_System.MEMCMP(ADR(vio_New), ADR(vo_Visu.stConfig), SIZEOF(vio_New)) <> 0;
IF m_ApplyConfig THEN
	vo_Visu.stConfig := vio_New;
	m_NotifyConfigChanged();
END_IF
END_METHOD

(****************************************************************************************************<br>
© Syntegon Group.<br>
All rights reserved, also regarding any disposal, exploitation, reproduction, editing, distribution,<br>
as well as in the event of applications for industrial property rights.<br>
*****************************************************************************************************<br>
DESCRIPTION:<br>
Belt position last set, [mm].<br>
****************************************************************************************************)
METHOD m_BeltPosition : LREAL
m_BeltPosition := vo_Visu.stState.fBeltPosition;
END_METHOD

(****************************************************************************************************<br>
© Syntegon Group.<br>
All rights reserved, also regarding any disposal, exploitation, reproduction, editing, distribution,<br>
as well as in the event of applications for industrial property rights.<br>
*****************************************************************************************************<br>
DESCRIPTION:<br>
Manifest type: conveyor.<br>
****************************************************************************************************)
METHOD PROTECTED m_ComponentType : E_VisuComponentType
m_ComponentType := E_VisuComponentType.CONVEYOR;
END_METHOD

(****************************************************************************************************<br>
© Syntegon Group.<br>
All rights reserved, also regarding any disposal, exploitation, reproduction, editing, distribution,<br>
as well as in the event of applications for industrial property rights.<br>
*****************************************************************************************************<br>
DESCRIPTION:<br>
Sets pose and size. TRUE if anything changed.<br>
****************************************************************************************************)
METHOD m_Configure : BOOL
VAR_INPUT
	vi_Pose								: ST_VisuPose;	// MCS, belt start on the belt surface; local +X = conveying direction
	vi_lr_Length						: LREAL;	// [mm]
	vi_lr_Width							: LREAL;	// [mm]
END_VAR
VAR
	TempNew								: ST_VisuConveyorConfig;
END_VAR
TempNew := vo_Visu.stConfig;
TempNew.stPose := vi_Pose;
TempNew.fLength := vi_lr_Length;
TempNew.fWidth := vi_lr_Width;
m_Configure := m_ApplyConfig(TempNew);
END_METHOD

(****************************************************************************************************<br>
© Syntegon Group.<br>
All rights reserved, also regarding any disposal, exploitation, reproduction, editing, distribution,<br>
as well as in the event of applications for industrial property rights.<br>
*****************************************************************************************************<br>
DESCRIPTION:<br>
Register index of the product with vi_udn_Id, -1 if not found.<br>
****************************************************************************************************)
METHOD m_FindProduct : INT
VAR_INPUT
	vi_udn_Id							: UDINT;	// [-] product id
END_VAR
VAR
	un_TempIndex						: UINT;
END_VAR
m_FindProduct := -1;
un_TempIndex := 0;
WHILE un_TempIndex < vo_Visu.stState.nProductCount DO
	IF vo_Visu.stState.aProducts[un_TempIndex].nId = vi_udn_Id THEN
		m_FindProduct := UINT_TO_INT(un_TempIndex);
		RETURN;
	END_IF
	un_TempIndex := un_TempIndex + 1;
END_WHILE
END_METHOD

(****************************************************************************************************<br>
© Syntegon Group.<br>
All rights reserved, also regarding any disposal, exploitation, reproduction, editing, distribution,<br>
as well as in the event of applications for industrial property rights.<br>
*****************************************************************************************************<br>
DESCRIPTION:<br>
Reads register entry vi_un_Index and its current MCS pose (latch pose moved by the belt travel since).<br>
Indices shift when products are removed; use the product id to follow a product.<br>
*****************************************************************************************************<br>
OUTPUT VALUES:<br>
FALSE if vi_un_Index is out of range.<br>
****************************************************************************************************)
METHOD m_GetProduct : BOOL
VAR_INPUT
	vi_un_Index							: UINT;	// [-] 0..m_ProductCount() - 1
END_VAR
VAR_OUTPUT
	vo_Product							: ST_VisuProduct;
	vo_Pose								: ST_VisuPlanarPose;	// MCS, current bottom centre
END_VAR
m_GetProduct := vi_un_Index < vo_Visu.stState.nProductCount;
IF m_GetProduct THEN
	vo_Product := vo_Visu.stState.aProducts[vi_un_Index];
	vo_Pose := m_ProductPose(vo_Product);
END_IF
END_METHOD

(****************************************************************************************************<br>
© Syntegon Group.<br>
All rights reserved, also regarding any disposal, exploitation, reproduction, editing, distribution,<br>
as well as in the event of applications for industrial property rights.<br>
*****************************************************************************************************<br>
DESCRIPTION:<br>
Adds a detected product at the current belt position. Call m_SetBeltPosition first in the cycle,<br>
or pass the belt position at the latch moment in vi_lr_LatchBeltPosition.<br>
*****************************************************************************************************<br>
OUTPUT VALUES:<br>
FALSE for vi_udn_Id = 0, an id already in the register, or a full register.<br>
****************************************************************************************************)
METHOD m_LatchProduct : BOOL
VAR_INPUT
	vi_udn_Id							: UDINT;	// [-] unique on this conveyor, > 0
	vi_LatchPose						: ST_VisuPlanarPose;	// MCS, bottom centre of the product at the latch moment
	vi_udn_ProductType					: UDINT;	// [-] id given to m_SetProductType
	vi_lr_LatchBeltPosition				: LREAL := 0;	// [mm] used only if vi_b_UseLatchBeltPosition
	vi_b_UseLatchBeltPosition			: BOOL := FALSE;	// FALSE: latch at the current belt position
END_VAR
VAR
	un_TempIndex						: UINT;
END_VAR
m_LatchProduct := FALSE;
un_TempIndex := vo_Visu.stState.nProductCount;
IF vi_udn_Id = 0 OR m_FindProduct(vi_udn_Id) >= 0 OR un_TempIndex >= VISU_GlobalConst_Param.VISU_un_MAX_PRODUCTS THEN
	RETURN;
END_IF
vo_Visu.stState.aProducts[un_TempIndex].nId := vi_udn_Id;
vo_Visu.stState.aProducts[un_TempIndex].bValid := TRUE;
vo_Visu.stState.aProducts[un_TempIndex].stLatchPose := vi_LatchPose;
IF vi_b_UseLatchBeltPosition THEN
	vo_Visu.stState.aProducts[un_TempIndex].fLatchBeltPosition := vi_lr_LatchBeltPosition;
ELSE
	vo_Visu.stState.aProducts[un_TempIndex].fLatchBeltPosition := vo_Visu.stState.fBeltPosition;
END_IF
vo_Visu.stState.aProducts[un_TempIndex].eState := E_VisuProductState.DETECTED;
vo_Visu.stState.aProducts[un_TempIndex].nRobotId := 0;
vo_Visu.stState.aProducts[un_TempIndex].nMoverId := 0;
vo_Visu.stState.aProducts[un_TempIndex].nProductType := vi_udn_ProductType;
vo_Visu.stState.nProductCount := un_TempIndex + 1;
vo_Visu.stState.nTimestamp := m_DcTime();
m_LatchProduct := TRUE;
END_METHOD

(****************************************************************************************************<br>
© Syntegon Group.<br>
All rights reserved, also regarding any disposal, exploitation, reproduction, editing, distribution,<br>
as well as in the event of applications for industrial property rights.<br>
*****************************************************************************************************<br>
DESCRIPTION:<br>
Puts a product of the register at a new MCS pose at the current belt position, e.g. while a mover pushes it<br>
along the belt faster than the belt runs. Call m_SetBeltPosition first in the cycle. Keeps its state.<br>
*****************************************************************************************************<br>
OUTPUT VALUES:<br>
FALSE if the product is not in the register.<br>
****************************************************************************************************)
METHOD m_MoveProduct : BOOL
VAR_INPUT
	vi_udn_Id							: UDINT;	// [-] product id
	vi_Pose								: ST_VisuPlanarPose;	// MCS, bottom centre of the product now
END_VAR
VAR
	n_TempIndex							: INT;
END_VAR
n_TempIndex := m_FindProduct(vi_udn_Id);
m_MoveProduct := n_TempIndex >= 0;
IF m_MoveProduct THEN
	vo_Visu.stState.aProducts[n_TempIndex].stLatchPose := vi_Pose;
	vo_Visu.stState.aProducts[n_TempIndex].fLatchBeltPosition := vo_Visu.stState.fBeltPosition;
	vo_Visu.stState.nTimestamp := m_DcTime();
END_IF
END_METHOD

(****************************************************************************************************<br>
© Syntegon Group.<br>
All rights reserved, also regarding any disposal, exploitation, reproduction, editing, distribution,<br>
as well as in the event of applications for industrial property rights.<br>
*****************************************************************************************************<br>
DESCRIPTION:<br>
Number of products in the register; valid indices for m_GetProduct are 0..m_ProductCount() - 1.<br>
****************************************************************************************************)
METHOD m_ProductCount : UINT
m_ProductCount := vo_Visu.stState.nProductCount;
END_METHOD

(****************************************************************************************************<br>
© Syntegon Group.<br>
All rights reserved, also regarding any disposal, exploitation, reproduction, editing, distribution,<br>
as well as in the event of applications for industrial property rights.<br>
*****************************************************************************************************<br>
DESCRIPTION:<br>
Current MCS pose of a product: latch pose moved along the conveying direction (local +X,<br>
rotation Rz * Ry of the conveyor pose) by the belt travel since the latch.<br>
****************************************************************************************************)
METHOD PRIVATE m_ProductPose : ST_VisuPlanarPose
VAR_IN_OUT CONSTANT
	vio_Product							: ST_VisuProduct;
END_VAR
VAR
	lr_TempTravel						: LREAL;	// [mm]
	lr_TempRz							: LREAL;	// [rad]
	lr_TempRy							: LREAL;	// [rad]
END_VAR
lr_TempTravel := vo_Visu.stState.fBeltPosition - vio_Product.fLatchBeltPosition;
lr_TempRz := vo_Visu.stConfig.stPose.fRz * VISU_GlobalConst.VISU_lr_DEG_TO_RAD;
lr_TempRy := vo_Visu.stConfig.stPose.fRy * VISU_GlobalConst.VISU_lr_DEG_TO_RAD;
m_ProductPose := vio_Product.stLatchPose;
m_ProductPose.fX := m_ProductPose.fX + lr_TempTravel * COS(lr_TempRz) * COS(lr_TempRy);
m_ProductPose.fY := m_ProductPose.fY + lr_TempTravel * SIN(lr_TempRz) * COS(lr_TempRy);
m_ProductPose.fZ := m_ProductPose.fZ - lr_TempTravel * SIN(lr_TempRy);
END_METHOD

(****************************************************************************************************<br>
© Syntegon Group.<br>
All rights reserved, also regarding any disposal, exploitation, reproduction, editing, distribution,<br>
as well as in the event of applications for industrial property rights.<br>
*****************************************************************************************************<br>
DESCRIPTION:<br>
Removes a product from the register. FALSE if it is not in the register.<br>
****************************************************************************************************)
METHOD m_RemoveProduct : BOOL
VAR_INPUT
	vi_udn_Id							: UDINT;	// [-] product id
END_VAR
VAR
	n_TempIndex							: INT;
	n_TempLast							: INT;
END_VAR
n_TempIndex := m_FindProduct(vi_udn_Id);
m_RemoveProduct := n_TempIndex >= 0;
IF NOT m_RemoveProduct THEN
	RETURN;
END_IF
n_TempLast := UINT_TO_INT(vo_Visu.stState.nProductCount) - 1;
WHILE n_TempIndex < n_TempLast DO
	vo_Visu.stState.aProducts[n_TempIndex] := vo_Visu.stState.aProducts[n_TempIndex + 1];
	n_TempIndex := n_TempIndex + 1;
END_WHILE
vo_Visu.stState.aProducts[n_TempLast].bValid := FALSE;
vo_Visu.stState.nProductCount := INT_TO_UINT(n_TempLast);
vo_Visu.stState.nTimestamp := m_DcTime();
END_METHOD

(****************************************************************************************************<br>
© Syntegon Group.<br>
All rights reserved, also regarding any disposal, exploitation, reproduction, editing, distribution,<br>
as well as in the event of applications for industrial property rights.<br>
*****************************************************************************************************<br>
DESCRIPTION:<br>
Housekeeping: drops invalid entries and products that have travelled beyond vi_lr_BeltX (along the<br>
conveyor from its start). Products a robot is working on (ASSIGNED or PICKED) are kept wherever they are.<br>
*****************************************************************************************************<br>
OUTPUT VALUES:<br>
Number of removed entries.<br>
****************************************************************************************************)
METHOD m_RemoveProductsBeyond : UINT
VAR_INPUT
	vi_lr_BeltX							: LREAL;	// [mm] e.g. belt length + some margin so missed products stay visible briefly
END_VAR
VAR
	un_TempRead							: UINT;
	un_TempWrite						: UINT;
	b_TempInUse							: BOOL;
	TempPose							: ST_VisuPlanarPose;
	lr_TempDx							: LREAL;	// [mm]
	lr_TempDy							: LREAL;	// [mm]
	lr_TempDz							: LREAL;	// [mm]
	lr_TempRz							: LREAL;	// [rad]
	lr_TempRy							: LREAL;	// [rad]
	lr_TempX							: LREAL;	// [mm] belt X
END_VAR
m_RemoveProductsBeyond := 0;
IF vo_Visu.stState.nProductCount = 0 THEN
	RETURN;
END_IF
lr_TempRz := vo_Visu.stConfig.stPose.fRz * VISU_GlobalConst.VISU_lr_DEG_TO_RAD;
lr_TempRy := vo_Visu.stConfig.stPose.fRy * VISU_GlobalConst.VISU_lr_DEG_TO_RAD;

(* Keep the entries to stay, in order. *)
un_TempWrite := 0;
FOR un_TempRead := 0 TO vo_Visu.stState.nProductCount - 1 DO
	(* Belt X = current position projected onto the conveying direction, measured from the belt start. *)
	TempPose := m_ProductPose(vo_Visu.stState.aProducts[un_TempRead]);
	lr_TempDx := TempPose.fX - vo_Visu.stConfig.stPose.fX;
	lr_TempDy := TempPose.fY - vo_Visu.stConfig.stPose.fY;
	lr_TempDz := TempPose.fZ - vo_Visu.stConfig.stPose.fZ;
	lr_TempX := (lr_TempDx * COS(lr_TempRz) + lr_TempDy * SIN(lr_TempRz)) * COS(lr_TempRy)
				- lr_TempDz * SIN(lr_TempRy);
	b_TempInUse := vo_Visu.stState.aProducts[un_TempRead].eState = E_VisuProductState.ASSIGNED
				OR vo_Visu.stState.aProducts[un_TempRead].eState = E_VisuProductState.PICKED;
	IF vo_Visu.stState.aProducts[un_TempRead].bValid AND (lr_TempX <= vi_lr_BeltX OR b_TempInUse) THEN
		IF un_TempWrite <> un_TempRead THEN
			vo_Visu.stState.aProducts[un_TempWrite] := vo_Visu.stState.aProducts[un_TempRead];
		END_IF
		un_TempWrite := un_TempWrite + 1;
	END_IF
END_FOR

(* Invalidate the freed tail. *)
m_RemoveProductsBeyond := vo_Visu.stState.nProductCount - un_TempWrite;
IF un_TempWrite < vo_Visu.stState.nProductCount THEN
	FOR un_TempRead := un_TempWrite TO vo_Visu.stState.nProductCount - 1 DO
		vo_Visu.stState.aProducts[un_TempRead].bValid := FALSE;
	END_FOR
	vo_Visu.stState.nProductCount := un_TempWrite;
	vo_Visu.stState.nTimestamp := m_DcTime();
END_IF
END_METHOD

(****************************************************************************************************<br>
© Syntegon Group.<br>
All rights reserved, also regarding any disposal, exploitation, reproduction, editing, distribution,<br>
as well as in the event of applications for industrial property rights.<br>
*****************************************************************************************************<br>
DESCRIPTION:<br>
Sets the belt position: how far the belt surface has travelled, continuous (no modulo).<br>
Call once per cycle; it also stamps the state with the cycle's DC time.<br>
****************************************************************************************************)
METHOD m_SetBeltPosition : BOOL
VAR_INPUT
	vi_lr_Position						: LREAL;	// [mm]
END_VAR
vo_Visu.stState.fBeltPosition := vi_lr_Position;
vo_Visu.stState.nTimestamp := m_DcTime();
m_SetBeltPosition := TRUE;
END_METHOD

(****************************************************************************************************<br>
© Syntegon Group.<br>
All rights reserved, also regarding any disposal, exploitation, reproduction, editing, distribution,<br>
as well as in the event of applications for industrial property rights.<br>
*****************************************************************************************************<br>
DESCRIPTION:<br>
Sets or clears the fault of the conveyor: drawn red with the message while active. The fault stays until it<br>
is cleared with m_SetFault(vi_b_Active := FALSE, vi_str_Message := ''). TRUE.<br>
****************************************************************************************************)
METHOD m_SetFault : BOOL
VAR_INPUT
	vi_b_Active							: BOOL;	// TRUE: fault active
	vi_str_Message						: STRING(80);	// shown to the operator; empty shows 'Fault'
END_VAR
vo_Visu.stState.stFault.bActive := vi_b_Active;
vo_Visu.stState.stFault.sMessage := vi_str_Message;
m_SetFault := TRUE;
END_METHOD

(****************************************************************************************************<br>
© Syntegon Group.<br>
All rights reserved, also regarding any disposal, exploitation, reproduction, editing, distribution,<br>
as well as in the event of applications for industrial property rights.<br>
*****************************************************************************************************<br>
DESCRIPTION:<br>
Like m_SetBeltPosition, for a modulo axis: unwraps the position so the belt position stays continuous.<br>
Call once per cycle.<br>
*****************************************************************************************************<br>
LIMITS:<br>
The axis must move less than half a modulo period per cycle.<br>
****************************************************************************************************)
METHOD m_SetModuloBeltPosition : BOOL
VAR_INPUT
	vi_lr_ModuloPosition				: LREAL;	// [mm] in [0, vi_lr_ModuloPeriod)
	vi_lr_ModuloPeriod					: LREAL;	// [mm] <= 0 passes vi_lr_ModuloPosition through unchanged
	vi_b_Reset							: BOOL;	// TRUE: restart the belt position at vi_lr_ModuloPosition
END_VAR
VAR
	lr_TempPosition						: LREAL;	// [mm]
	lr_TempDelta						: LREAL;	// [mm]
END_VAR
IF vi_b_Reset OR NOT b_ModuloInitialised OR vi_lr_ModuloPeriod <= 0 THEN
	lr_TempPosition := vi_lr_ModuloPosition;
	b_ModuloInitialised := TRUE;
ELSE
	lr_TempDelta := vi_lr_ModuloPosition - lr_LastModuloPosition;
	IF lr_TempDelta > vi_lr_ModuloPeriod / 2 THEN
		lr_TempDelta := lr_TempDelta - vi_lr_ModuloPeriod;
	ELSIF lr_TempDelta < -vi_lr_ModuloPeriod / 2 THEN
		lr_TempDelta := lr_TempDelta + vi_lr_ModuloPeriod;
	END_IF
	lr_TempPosition := vo_Visu.stState.fBeltPosition + lr_TempDelta;
END_IF
lr_LastModuloPosition := vi_lr_ModuloPosition;
m_SetModuloBeltPosition := m_SetBeltPosition(lr_TempPosition);
END_METHOD

(****************************************************************************************************<br>
© Syntegon Group.<br>
All rights reserved, also regarding any disposal, exploitation, reproduction, editing, distribution,<br>
as well as in the event of applications for industrial property rights.<br>
*****************************************************************************************************<br>
DESCRIPTION:<br>
Changes a product's state and assigned robot. FALSE if the product is not in the register.<br>
****************************************************************************************************)
METHOD m_SetProductState : BOOL
VAR_INPUT
	vi_udn_Id							: UDINT;	// [-] product id
	vi_e_State							: E_VisuProductState;
	vi_udn_RobotId						: UDINT;	// [-] manifest id of the robot, 0 = none
	vi_udn_MoverId						: UDINT := 0;	// [-] mover of an XTS gantry or loop carrying the product, 0 = none
	vi_udn_FingerId						: UDINT := 0;	// [-] gripper finger (1-based) the product hangs from while picked, 0 = the flange
END_VAR
VAR
	n_TempIndex							: INT;
END_VAR
n_TempIndex := m_FindProduct(vi_udn_Id);
m_SetProductState := n_TempIndex >= 0;
IF m_SetProductState THEN
	vo_Visu.stState.aProducts[n_TempIndex].eState := vi_e_State;
	vo_Visu.stState.aProducts[n_TempIndex].nRobotId := vi_udn_RobotId;
	vo_Visu.stState.aProducts[n_TempIndex].nMoverId := vi_udn_MoverId;
	vo_Visu.stState.aProducts[n_TempIndex].nFingerId := vi_udn_FingerId;
	vo_Visu.stState.nTimestamp := m_DcTime();
END_IF
END_METHOD

(****************************************************************************************************<br>
© Syntegon Group.<br>
All rights reserved, also regarding any disposal, exploitation, reproduction, editing, distribution,<br>
as well as in the event of applications for industrial property rights.<br>
*****************************************************************************************************<br>
DESCRIPTION:<br>
Adds a product type, or updates the one with the same id. FALSE for vi_udn_Id = 0 or a full list.<br>
****************************************************************************************************)
METHOD m_SetProductType : BOOL
VAR_INPUT
	vi_udn_Id							: UDINT;	// [-] referenced by m_LatchProduct's vi_udn_ProductType
	vi_lr_Length						: LREAL;	// [mm] along the conveying direction
	vi_lr_Width							: LREAL;	// [mm]
	vi_lr_Height						: LREAL;	// [mm]
END_VAR
VAR
	TempNew								: ST_VisuConveyorConfig;
	un_TempIndex						: UINT;
END_VAR
m_SetProductType := FALSE;
IF vi_udn_Id = 0 THEN
	RETURN;
END_IF
TempNew := vo_Visu.stConfig;
un_TempIndex := 0;
(* ST evaluates both operands of AND: test the index before reading the array. *)
WHILE un_TempIndex < TempNew.nProductTypeCount DO
	IF TempNew.aProductTypes[un_TempIndex].nId = vi_udn_Id THEN
		EXIT;
	END_IF
	un_TempIndex := un_TempIndex + 1;
END_WHILE
IF un_TempIndex >= VISU_GlobalConst_Param.VISU_un_MAX_PRODUCT_TYPES THEN
	RETURN;
END_IF
IF un_TempIndex = TempNew.nProductTypeCount THEN
	TempNew.nProductTypeCount := TempNew.nProductTypeCount + 1;
END_IF
TempNew.aProductTypes[un_TempIndex].nId := vi_udn_Id;
TempNew.aProductTypes[un_TempIndex].fLength := vi_lr_Length;
TempNew.aProductTypes[un_TempIndex].fWidth := vi_lr_Width;
TempNew.aProductTypes[un_TempIndex].fHeight := vi_lr_Height;
m_ApplyConfig(TempNew);
m_SetProductType := TRUE;
END_METHOD

END_FUNCTION_BLOCK

// POUs/_FB_VisuDelta
(****************************************************************************************************<br>
© Syntegon Group.<br>
All rights reserved, also regarding any disposal, exploitation, reproduction, editing, distribution,<br>
as well as in the event of applications for industrial property rights.<br>
*****************************************************************************************************<br>
DESCRIPTION:<br>
One visualised Delta robot. Typical cycle:<br>
  fb_Delta.m_Register(vio_Manifest := GVL_Visu.stManifest, vi_udn_Id := 10, vi_str_Name := 'Delta 1',<br>
      vi_str_Path := 'MAIN.fb_Delta.vo_Visu');<br>
  fb_Delta.m_Configure(vi_Pose := BasePose, vi_lr_BaseRadius := 200, vi_lr_EffectorRadius := 50,<br>
      vi_lr_UpperArmLength := 400, vi_lr_LowerArmLength := 1000);<br>
  fb_Delta.m_SetFinger(vi_un_Finger := 1, vi_lr_Diameter := 40, vi_lr_Height := 50);<br>
  fb_Delta.m_SetWorkingArea(vi_lr_Radius := 750, vi_lr_ZMin := -1300, vi_lr_ZMax := -700, vi_lr_ConeHeight := 200,<br>
      vi_lr_ConeBottomRadius := 450);<br>
  fb_Delta.m_SetLimitArea(vi_lr_XMin := -500, vi_lr_XMax := 500, vi_lr_YMin := -750, vi_lr_YMax := 750,<br>
      vi_lr_ZMin := -1500, vi_lr_ZMax := -700);<br>
  fb_Delta.m_SetZone(vi_udn_ConveyorId := 1, vi_e_Kind := E_VisuZoneKind.PICK, vi_lr_Start := 1100, vi_lr_End := 1900,<br>
      vi_lr_AllocationOffset := 300);<br>
  fb_Delta.m_SetTcp(vi_ActualTcp := ActualTcp, vi_SetpointTcp := SetpointTcp);<br>
  fb_Delta.m_SetFingerState(vi_un_Finger := 1, vi_Pose := CupPose, vi_b_Active := b_Vacuum);<br>
Only the TCP (the gripper flange) is reported; the visualisation derives the arms from it. Tool rotations<br>
(e.g. a 4th axis) show only through the finger poses, absolute in the MCS. The config methods may be called<br>
every cycle; the config version only changes when a value does.<br>
*****************************************************************************************************<br>
OUTPUT VALUES:<br>
vo_Visu is the contract structure the gateway reads at the path given to m_Register. Do not write it.<br>
*****************************************************************************************************<br>
VERSION         ¦ DATE       ¦ NAME      ¦ CHANGE<br>
Syn_Visu 3.0.0  ¦ 2026-10-31 ¦ J.Willner ¦ Naming and layout after the TCAT programming guideline<br>
****************************************************************************************************)
FUNCTION_BLOCK _FB_VisuDelta EXTENDS _FB_VisuComponent
VAR_OUTPUT
	vo_Visu								: ST_VisuDelta;	// contract structure read by the gateway
END_VAR

(****************************************************************************************************<br>
© Syntegon Group.<br>
All rights reserved, also regarding any disposal, exploitation, reproduction, editing, distribution,<br>
as well as in the event of applications for industrial property rights.<br>
*****************************************************************************************************<br>
DESCRIPTION:<br>
Takes over vio_New and increments the config version if it differs from the current config. TRUE if changed.<br>
****************************************************************************************************)
METHOD PRIVATE m_ApplyConfig : BOOL
VAR_IN_OUT
	vio_New								: ST_VisuDeltaConfig;
END_VAR
m_ApplyConfig := Tc2_System.MEMCMP(ADR(vio_New), ADR(vo_Visu.stConfig), SIZEOF(vio_New)) <> 0;
IF m_ApplyConfig THEN
	vo_Visu.stConfig := vio_New;
	m_NotifyConfigChanged();
END_IF
END_METHOD

(****************************************************************************************************<br>
© Syntegon Group.<br>
All rights reserved, also regarding any disposal, exploitation, reproduction, editing, distribution,<br>
as well as in the event of applications for industrial property rights.<br>
*****************************************************************************************************<br>
DESCRIPTION:<br>
Base pose last set by m_Configure, MCS.<br>
****************************************************************************************************)
METHOD m_BasePose : ST_VisuPose
m_BasePose := vo_Visu.stConfig.stPose;
END_METHOD

(****************************************************************************************************<br>
© Syntegon Group.<br>
All rights reserved, also regarding any disposal, exploitation, reproduction, editing, distribution,<br>
as well as in the event of applications for industrial property rights.<br>
*****************************************************************************************************<br>
DESCRIPTION:<br>
Removes the gripper definition. TRUE if there was one.<br>
****************************************************************************************************)
METHOD m_ClearFingers : BOOL
VAR
	TempNew								: ST_VisuDeltaConfig;
	TempEmpty							: ST_VisuFinger;
	un_TempIndex						: UINT;
END_VAR
TempNew := vo_Visu.stConfig;
FOR un_TempIndex := 0 TO VISU_GlobalConst_Param.VISU_un_MAX_FINGERS - 1 DO
	TempNew.aFingers[un_TempIndex] := TempEmpty;
END_FOR
TempNew.nFingerCount := 0;
m_ClearFingers := m_ApplyConfig(TempNew);
END_METHOD

(****************************************************************************************************<br>
© Syntegon Group.<br>
All rights reserved, also regarding any disposal, exploitation, reproduction, editing, distribution,<br>
as well as in the event of applications for industrial property rights.<br>
*****************************************************************************************************<br>
DESCRIPTION:<br>
Removes the limit area. TRUE if changed.<br>
****************************************************************************************************)
METHOD m_ClearLimitArea : BOOL
VAR
	TempNew								: ST_VisuDeltaConfig;
	TempEmpty							: ST_VisuLimitArea;
END_VAR
TempNew := vo_Visu.stConfig;
TempNew.stLimitArea := TempEmpty;
m_ClearLimitArea := m_ApplyConfig(TempNew);
END_METHOD

(****************************************************************************************************<br>
© Syntegon Group.<br>
All rights reserved, also regarding any disposal, exploitation, reproduction, editing, distribution,<br>
as well as in the event of applications for industrial property rights.<br>
*****************************************************************************************************<br>
DESCRIPTION:<br>
Removes all pick and place zones. TRUE if there were any.<br>
****************************************************************************************************)
METHOD m_ClearZones : BOOL
VAR
	TempNew								: ST_VisuDeltaConfig;
	TempEmpty							: ST_VisuZone;
	un_TempIndex						: UINT;
END_VAR
TempNew := vo_Visu.stConfig;
FOR un_TempIndex := 0 TO VISU_GlobalConst_Param.VISU_un_MAX_ZONES - 1 DO
	TempNew.aZones[un_TempIndex] := TempEmpty;
END_FOR
TempNew.nZoneCount := 0;
m_ClearZones := m_ApplyConfig(TempNew);
END_METHOD

(****************************************************************************************************<br>
© Syntegon Group.<br>
All rights reserved, also regarding any disposal, exploitation, reproduction, editing, distribution,<br>
as well as in the event of applications for industrial property rights.<br>
*****************************************************************************************************<br>
DESCRIPTION:<br>
Manifest type: Delta robot.<br>
****************************************************************************************************)
METHOD PROTECTED m_ComponentType : E_VisuComponentType
m_ComponentType := E_VisuComponentType.DELTA;
END_METHOD

(****************************************************************************************************<br>
© Syntegon Group.<br>
All rights reserved, also regarding any disposal, exploitation, reproduction, editing, distribution,<br>
as well as in the event of applications for industrial property rights.<br>
*****************************************************************************************************<br>
DESCRIPTION:<br>
Sets base pose and geometry. Arm 1 lies along the base's local +X; arms 2 and 3 follow<br>
counter-clockwise (seen from above) at 120 deg each. TRUE if anything changed.<br>
****************************************************************************************************)
METHOD m_Configure : BOOL
VAR_INPUT
	vi_Pose								: ST_VisuPose;	// MCS, base centre
	vi_lr_BaseRadius					: LREAL;	// [mm] base centre to shoulder joint
	vi_lr_EffectorRadius				: LREAL;	// [mm] effector centre to lower-arm joint
	vi_lr_UpperArmLength				: LREAL;	// [mm]
	vi_lr_LowerArmLength				: LREAL;	// [mm]
END_VAR
VAR
	TempNew								: ST_VisuDeltaConfig;
END_VAR
TempNew := vo_Visu.stConfig;
TempNew.stPose := vi_Pose;
TempNew.fBaseRadius := vi_lr_BaseRadius;
TempNew.fEffectorRadius := vi_lr_EffectorRadius;
TempNew.fUpperArmLength := vi_lr_UpperArmLength;
TempNew.fLowerArmLength := vi_lr_LowerArmLength;
m_Configure := m_ApplyConfig(TempNew);
END_METHOD

(****************************************************************************************************<br>
© Syntegon Group.<br>
All rights reserved, also regarding any disposal, exploitation, reproduction, editing, distribution,<br>
as well as in the event of applications for industrial property rights.<br>
*****************************************************************************************************<br>
DESCRIPTION:<br>
Sets or clears the fault of the robot: drawn red with the message while active. The fault stays until it<br>
is cleared with m_SetFault(vi_b_Active := FALSE, vi_str_Message := ''). TRUE.<br>
****************************************************************************************************)
METHOD m_SetFault : BOOL
VAR_INPUT
	vi_b_Active							: BOOL;	// TRUE: fault active
	vi_str_Message						: STRING(80);	// shown to the operator; empty shows 'Fault'
END_VAR
vo_Visu.stState.stFault.bActive := vi_b_Active;
vo_Visu.stState.stFault.sMessage := vi_str_Message;
m_SetFault := TRUE;
END_METHOD

(****************************************************************************************************<br>
© Syntegon Group.<br>
All rights reserved, also regarding any disposal, exploitation, reproduction, editing, distribution,<br>
as well as in the event of applications for industrial property rights.<br>
*****************************************************************************************************<br>
DESCRIPTION:<br>
Defines gripper finger vi_un_Finger (1-based): a cylinder hanging from the finger's pose along its local -Z.<br>
The finger count grows to vi_un_Finger.<br>
*****************************************************************************************************<br>
OUTPUT VALUES:<br>
FALSE outside 1..VISU_GlobalConst_Param.VISU_un_MAX_FINGERS.<br>
****************************************************************************************************)
METHOD m_SetFinger : BOOL
VAR_INPUT
	vi_un_Finger						: UINT;	// [-] 1-based, as a product's nFingerId
	vi_lr_Diameter						: LREAL;	// [mm]
	vi_lr_Height						: LREAL;	// [mm] along the finger's local -Z
END_VAR
VAR
	TempNew								: ST_VisuDeltaConfig;
END_VAR
m_SetFinger := FALSE;
IF vi_un_Finger = 0 OR vi_un_Finger > VISU_GlobalConst_Param.VISU_un_MAX_FINGERS THEN
	RETURN;
END_IF
TempNew := vo_Visu.stConfig;
TempNew.aFingers[vi_un_Finger - 1].fDiameter := vi_lr_Diameter;
TempNew.aFingers[vi_un_Finger - 1].fHeight := vi_lr_Height;
TempNew.nFingerCount := MAX(TempNew.nFingerCount, vi_un_Finger);
m_ApplyConfig(TempNew);
m_SetFinger := TRUE;
END_METHOD

(****************************************************************************************************<br>
© Syntegon Group.<br>
All rights reserved, also regarding any disposal, exploitation, reproduction, editing, distribution,<br>
as well as in the event of applications for industrial property rights.<br>
*****************************************************************************************************<br>
DESCRIPTION:<br>
Reports finger vi_un_Finger (1-based): the pose of its frame (centre of its top face), absolute in the MCS,<br>
and whether it grips. Call once per cycle per configured finger.<br>
*****************************************************************************************************<br>
OUTPUT VALUES:<br>
FALSE outside 1..VISU_GlobalConst_Param.VISU_un_MAX_FINGERS.<br>
****************************************************************************************************)
METHOD m_SetFingerState : BOOL
VAR_INPUT
	vi_un_Finger						: UINT;	// [-] 1-based
	vi_Pose								: ST_VisuPose;	// MCS
	vi_b_Active							: BOOL;	// TRUE while the finger grips
END_VAR
m_SetFingerState := vi_un_Finger > 0 AND vi_un_Finger <= VISU_GlobalConst_Param.VISU_un_MAX_FINGERS;
IF m_SetFingerState THEN
	vo_Visu.stState.aFingerStates[vi_un_Finger - 1].stPose := vi_Pose;
	vo_Visu.stState.aFingerStates[vi_un_Finger - 1].bActive := vi_b_Active;
END_IF
END_METHOD

(****************************************************************************************************<br>
© Syntegon Group.<br>
All rights reserved, also regarding any disposal, exploitation, reproduction, editing, distribution,<br>
as well as in the event of applications for industrial property rights.<br>
*****************************************************************************************************<br>
DESCRIPTION:<br>
Sets and activates the limit area: an axis-aligned box in the robot frame. TRUE if changed.<br>
****************************************************************************************************)
METHOD m_SetLimitArea : BOOL
VAR_INPUT
	vi_lr_XMin							: LREAL;	// [mm]
	vi_lr_XMax							: LREAL;	// [mm]
	vi_lr_YMin							: LREAL;	// [mm]
	vi_lr_YMax							: LREAL;	// [mm]
	vi_lr_ZMin							: LREAL;	// [mm] relative to the base (below the base: negative)
	vi_lr_ZMax							: LREAL;	// [mm] relative to the base
END_VAR
VAR
	TempNew								: ST_VisuDeltaConfig;
END_VAR
TempNew := vo_Visu.stConfig;
TempNew.stLimitArea.fXMin := vi_lr_XMin;
TempNew.stLimitArea.fXMax := vi_lr_XMax;
TempNew.stLimitArea.fYMin := vi_lr_YMin;
TempNew.stLimitArea.fYMax := vi_lr_YMax;
TempNew.stLimitArea.fZMin := vi_lr_ZMin;
TempNew.stLimitArea.fZMax := vi_lr_ZMax;
TempNew.stLimitArea.bActive := TRUE;
m_SetLimitArea := m_ApplyConfig(TempNew);
END_METHOD

(****************************************************************************************************<br>
© Syntegon Group.<br>
All rights reserved, also regarding any disposal, exploitation, reproduction, editing, distribution,<br>
as well as in the event of applications for industrial property rights.<br>
*****************************************************************************************************<br>
DESCRIPTION:<br>
Reports the robot's TCP. Call once per cycle; it also stamps the state with the cycle's DC time.<br>
****************************************************************************************************)
METHOD m_SetTcp : BOOL
VAR_INPUT
	vi_ActualTcp						: ST_VisuPosition;	// MCS, effector centre (the gripper flange)
	vi_SetpointTcp						: ST_VisuPosition;	// MCS
END_VAR
vo_Visu.stState.stActualTcp := vi_ActualTcp;
vo_Visu.stState.stSetpointTcp := vi_SetpointTcp;
vo_Visu.stState.nTimestamp := m_DcTime();
m_SetTcp := TRUE;
END_METHOD

(****************************************************************************************************<br>
© Syntegon Group.<br>
All rights reserved, also regarding any disposal, exploitation, reproduction, editing, distribution,<br>
as well as in the event of applications for industrial property rights.<br>
*****************************************************************************************************<br>
DESCRIPTION:<br>
Sets the working area: a vertical cylinder in the robot frame with an optional cone below. TRUE if changed.<br>
****************************************************************************************************)
METHOD m_SetWorkingArea : BOOL
VAR_INPUT
	vi_lr_Radius						: LREAL;	// [mm]
	vi_lr_ZMin							: LREAL;	// [mm] relative to the base (below the base: negative)
	vi_lr_ZMax							: LREAL;	// [mm] relative to the base
	vi_lr_ConeHeight					: LREAL;	// [mm] below vi_lr_ZMin; 0 = no cone
	vi_lr_ConeBottomRadius				: LREAL;	// [mm]
END_VAR
VAR
	TempNew								: ST_VisuDeltaConfig;
END_VAR
TempNew := vo_Visu.stConfig;
TempNew.stWorkingArea.fRadius := vi_lr_Radius;
TempNew.stWorkingArea.fZMin := vi_lr_ZMin;
TempNew.stWorkingArea.fZMax := vi_lr_ZMax;
TempNew.stWorkingArea.fConeHeight := vi_lr_ConeHeight;
TempNew.stWorkingArea.fConeBottomRadius := vi_lr_ConeBottomRadius;
m_SetWorkingArea := m_ApplyConfig(TempNew);
END_METHOD

(****************************************************************************************************<br>
© Syntegon Group.<br>
All rights reserved, also regarding any disposal, exploitation, reproduction, editing, distribution,<br>
as well as in the event of applications for industrial property rights.<br>
*****************************************************************************************************<br>
DESCRIPTION:<br>
Adds a pick or place zone, or updates the one for the same conveyor and kind.<br>
*****************************************************************************************************<br>
OUTPUT VALUES:<br>
FALSE for vi_udn_ConveyorId = 0 or a full list.<br>
****************************************************************************************************)
METHOD m_SetZone : BOOL
VAR_INPUT
	vi_udn_ConveyorId					: UDINT;	// [-] manifest id of the conveyor
	vi_e_Kind							: E_VisuZoneKind;
	vi_lr_Start							: LREAL;	// [mm] along the conveyor from its start (belt coordinates, not MCS)
	vi_lr_End							: LREAL;	// [mm] along the conveyor from its start
	vi_lr_AllocationOffset				: LREAL := 0;	// [mm] before vi_lr_End up to which products may be allocated; 0 = no limit
END_VAR
VAR
	TempNew								: ST_VisuDeltaConfig;
	un_TempIndex						: UINT;
END_VAR
m_SetZone := FALSE;
IF vi_udn_ConveyorId = 0 THEN
	RETURN;
END_IF
TempNew := vo_Visu.stConfig;
un_TempIndex := 0;
(* ST evaluates both operands of AND: test the index before reading the array. *)
WHILE un_TempIndex < TempNew.nZoneCount DO
	IF TempNew.aZones[un_TempIndex].nConveyorId = vi_udn_ConveyorId AND TempNew.aZones[un_TempIndex].eKind = vi_e_Kind THEN
		EXIT;
	END_IF
	un_TempIndex := un_TempIndex + 1;
END_WHILE
IF un_TempIndex >= VISU_GlobalConst_Param.VISU_un_MAX_ZONES THEN
	RETURN;
END_IF
IF un_TempIndex = TempNew.nZoneCount THEN
	TempNew.nZoneCount := TempNew.nZoneCount + 1;
END_IF
TempNew.aZones[un_TempIndex].nConveyorId := vi_udn_ConveyorId;
TempNew.aZones[un_TempIndex].eKind := vi_e_Kind;
TempNew.aZones[un_TempIndex].fStart := vi_lr_Start;
TempNew.aZones[un_TempIndex].fEnd := vi_lr_End;
TempNew.aZones[un_TempIndex].fAllocationOffset := vi_lr_AllocationOffset;
m_ApplyConfig(TempNew);
m_SetZone := TRUE;
END_METHOD

END_FUNCTION_BLOCK

// POUs/_FB_VisuXtsGantry
(****************************************************************************************************<br>
© Syntegon Group.<br>
All rights reserved, also regarding any disposal, exploitation, reproduction, editing, distribution,<br>
as well as in the event of applications for industrial property rights.<br>
*****************************************************************************************************<br>
DESCRIPTION:<br>
One visualised XTS gantry (e.g. IDH): a straight XTS track on a common Z axis, each mover with an X axis and a<br>
gripper flange at its end. Typical cycle:<br>
  fb_Idh.m_Register(vio_Manifest := GVL_Visu.stManifest, vi_udn_Id := 30, vi_str_Name := 'IDH',<br>
      vi_str_Path := 'MAIN.fb_Idh.vo_Visu');<br>
  fb_Idh.m_Configure(vi_Pose := TrackPose, vi_un_ModuleCount := 6, vi_lr_ModuleLength := 250, vi_lr_XMin := 0,<br>
      vi_lr_XMax := 700, vi_lr_ZMin := -100, vi_lr_ZMax := 0, vi_lr_ToolOffsetX := 150, vi_lr_ToolOffsetZ := -350,<br>
      vi_lr_MoverLength := 155, vi_lr_MoverWidth := 80);<br>
  fb_Idh.m_SetFinger(vi_un_Finger := 1, vi_lr_Diameter := 40, vi_lr_Height := 50);<br>
  fb_Idh.m_SetZone(vi_udn_ConveyorId := 3, vi_e_Kind := E_VisuZoneKind.PICK, vi_lr_Start := 1100, vi_lr_End := 2600);<br>
  fb_Idh.m_SetZPosition(lr_ZAxisActual);<br>
  fb_Idh.m_SetMoverCount(4);<br>
  fb_Idh.m_SetMover(vi_un_Index := 0, vi_udn_Id := 1, vi_lr_Position := ..., vi_lr_X := ..., vi_FingerStates := Mover1Fingers);<br>
Only actual values are reported; tool rotations (e.g. C) show only through the finger poses, absolute in the MCS.<br>
The config methods may be called every cycle; the config version only changes when a value does.<br>
*****************************************************************************************************<br>
OUTPUT VALUES:<br>
vo_Visu is the contract structure the gateway reads at the path given to m_Register. Do not write it.<br>
*****************************************************************************************************<br>
VERSION         ¦ DATE       ¦ NAME      ¦ CHANGE<br>
Syn_Visu 3.0.0  ¦ 2026-10-31 ¦ J.Willner ¦ Naming and layout after the TCAT programming guideline<br>
****************************************************************************************************)
FUNCTION_BLOCK _FB_VisuXtsGantry EXTENDS _FB_VisuComponent
VAR_OUTPUT
	vo_Visu								: ST_VisuXtsGantry;	// contract structure read by the gateway
END_VAR

(****************************************************************************************************<br>
© Syntegon Group.<br>
All rights reserved, also regarding any disposal, exploitation, reproduction, editing, distribution,<br>
as well as in the event of applications for industrial property rights.<br>
*****************************************************************************************************<br>
DESCRIPTION:<br>
Takes over vio_New and increments the config version if it differs from the current config. TRUE if changed.<br>
****************************************************************************************************)
METHOD PRIVATE m_ApplyConfig : BOOL
VAR_IN_OUT
	vio_New								: ST_VisuXtsGantryConfig;
END_VAR
m_ApplyConfig := Tc2_System.MEMCMP(ADR(vio_New), ADR(vo_Visu.stConfig), SIZEOF(vio_New)) <> 0;
IF m_ApplyConfig THEN
	vo_Visu.stConfig := vio_New;
	m_NotifyConfigChanged();
END_IF
END_METHOD

(****************************************************************************************************<br>
© Syntegon Group.<br>
All rights reserved, also regarding any disposal, exploitation, reproduction, editing, distribution,<br>
as well as in the event of applications for industrial property rights.<br>
*****************************************************************************************************<br>
DESCRIPTION:<br>
Removes the gripper definition. TRUE if there was one.<br>
****************************************************************************************************)
METHOD m_ClearFingers : BOOL
VAR
	TempNew								: ST_VisuXtsGantryConfig;
	TempEmpty							: ST_VisuFinger;
	un_TempIndex						: UINT;
END_VAR
TempNew := vo_Visu.stConfig;
FOR un_TempIndex := 0 TO VISU_GlobalConst_Param.VISU_un_MAX_FINGERS - 1 DO
	TempNew.aFingers[un_TempIndex] := TempEmpty;
END_FOR
TempNew.nFingerCount := 0;
m_ClearFingers := m_ApplyConfig(TempNew);
END_METHOD

(****************************************************************************************************<br>
© Syntegon Group.<br>
All rights reserved, also regarding any disposal, exploitation, reproduction, editing, distribution,<br>
as well as in the event of applications for industrial property rights.<br>
*****************************************************************************************************<br>
DESCRIPTION:<br>
Removes all pick and place zones. TRUE if there were any.<br>
****************************************************************************************************)
METHOD m_ClearZones : BOOL
VAR
	TempNew								: ST_VisuXtsGantryConfig;
	TempEmpty							: ST_VisuZone;
	un_TempIndex						: UINT;
END_VAR
TempNew := vo_Visu.stConfig;
FOR un_TempIndex := 0 TO VISU_GlobalConst_Param.VISU_un_MAX_ZONES - 1 DO
	TempNew.aZones[un_TempIndex] := TempEmpty;
END_FOR
TempNew.nZoneCount := 0;
m_ClearZones := m_ApplyConfig(TempNew);
END_METHOD

(****************************************************************************************************<br>
© Syntegon Group.<br>
All rights reserved, also regarding any disposal, exploitation, reproduction, editing, distribution,<br>
as well as in the event of applications for industrial property rights.<br>
*****************************************************************************************************<br>
DESCRIPTION:<br>
Manifest type: XTS gantry.<br>
****************************************************************************************************)
METHOD PROTECTED m_ComponentType : E_VisuComponentType
m_ComponentType := E_VisuComponentType.XTS_GANTRY;
END_METHOD

(****************************************************************************************************<br>
© Syntegon Group.<br>
All rights reserved, also regarding any disposal, exploitation, reproduction, editing, distribution,<br>
as well as in the event of applications for industrial property rights.<br>
*****************************************************************************************************<br>
DESCRIPTION:<br>
Sets pose, track, strokes, gripper offsets and mover size. TRUE if anything changed.<br>
****************************************************************************************************)
METHOD m_Configure : BOOL
VAR_INPUT
	vi_Pose								: ST_VisuPose;	// MCS, track start on top of the movers with Z = 0
	vi_un_ModuleCount					: UINT;	// [-] track modules in a row
	vi_lr_ModuleLength					: LREAL;	// [mm]
	vi_lr_XMin							: LREAL;	// [mm]
	vi_lr_XMax							: LREAL;	// [mm]
	vi_lr_ZMin							: LREAL;	// [mm]
	vi_lr_ZMax							: LREAL;	// [mm]
	vi_lr_ToolOffsetX					: LREAL;	// [mm] gripper flange ahead of the X axis zero
	vi_lr_ToolOffsetZ					: LREAL;	// [mm] gripper flange relative to the mover top (below: negative)
	vi_lr_MoverLength					: LREAL;	// [mm] along the track
	vi_lr_MoverWidth					: LREAL;	// [mm]
END_VAR
VAR
	TempNew								: ST_VisuXtsGantryConfig;
END_VAR
TempNew := vo_Visu.stConfig;
TempNew.stPose := vi_Pose;
TempNew.nModuleCount := vi_un_ModuleCount;
TempNew.fModuleLength := vi_lr_ModuleLength;
TempNew.fXMin := vi_lr_XMin;
TempNew.fXMax := vi_lr_XMax;
TempNew.fZMin := vi_lr_ZMin;
TempNew.fZMax := vi_lr_ZMax;
TempNew.fToolOffsetX := vi_lr_ToolOffsetX;
TempNew.fToolOffsetZ := vi_lr_ToolOffsetZ;
TempNew.fMoverLength := vi_lr_MoverLength;
TempNew.fMoverWidth := vi_lr_MoverWidth;
m_Configure := m_ApplyConfig(TempNew);
END_METHOD

(****************************************************************************************************<br>
© Syntegon Group.<br>
All rights reserved, also regarding any disposal, exploitation, reproduction, editing, distribution,<br>
as well as in the event of applications for industrial property rights.<br>
*****************************************************************************************************<br>
DESCRIPTION:<br>
Sets or clears the fault of the whole gantry: drawn red with the message while active. Faults of single<br>
movers go through m_SetMover. The fault stays until it is cleared with m_SetFault(vi_b_Active := FALSE,<br>
vi_str_Message := ''). TRUE.<br>
****************************************************************************************************)
METHOD m_SetFault : BOOL
VAR_INPUT
	vi_b_Active							: BOOL;	// TRUE: fault active
	vi_str_Message						: STRING(80);	// shown to the operator; empty shows 'Fault'
END_VAR
vo_Visu.stState.stFault.bActive := vi_b_Active;
vo_Visu.stState.stFault.sMessage := vi_str_Message;
m_SetFault := TRUE;
END_METHOD

(****************************************************************************************************<br>
© Syntegon Group.<br>
All rights reserved, also regarding any disposal, exploitation, reproduction, editing, distribution,<br>
as well as in the event of applications for industrial property rights.<br>
*****************************************************************************************************<br>
DESCRIPTION:<br>
Defines finger vi_un_Finger (1-based) of every mover's gripper: a cylinder hanging from the finger's pose along<br>
its local -Z. The finger count grows to vi_un_Finger.<br>
*****************************************************************************************************<br>
OUTPUT VALUES:<br>
FALSE outside 1..VISU_GlobalConst_Param.VISU_un_MAX_FINGERS.<br>
****************************************************************************************************)
METHOD m_SetFinger : BOOL
VAR_INPUT
	vi_un_Finger						: UINT;	// [-] 1-based, as a product's nFingerId
	vi_lr_Diameter						: LREAL;	// [mm]
	vi_lr_Height						: LREAL;	// [mm] along the finger's local -Z
END_VAR
VAR
	TempNew								: ST_VisuXtsGantryConfig;
END_VAR
m_SetFinger := FALSE;
IF vi_un_Finger = 0 OR vi_un_Finger > VISU_GlobalConst_Param.VISU_un_MAX_FINGERS THEN
	RETURN;
END_IF
TempNew := vo_Visu.stConfig;
TempNew.aFingers[vi_un_Finger - 1].fDiameter := vi_lr_Diameter;
TempNew.aFingers[vi_un_Finger - 1].fHeight := vi_lr_Height;
TempNew.nFingerCount := MAX(TempNew.nFingerCount, vi_un_Finger);
m_ApplyConfig(TempNew);
m_SetFinger := TRUE;
END_METHOD

(****************************************************************************************************<br>
© Syntegon Group.<br>
All rights reserved, also regarding any disposal, exploitation, reproduction, editing, distribution,<br>
as well as in the event of applications for industrial property rights.<br>
*****************************************************************************************************<br>
DESCRIPTION:<br>
Reports one mover (actual values) at entry vi_un_Index and marks it valid. Call once per cycle per mover.<br>
*****************************************************************************************************<br>
OUTPUT VALUES:<br>
FALSE if vi_un_Index is outside the mover count set by m_SetMoverCount.<br>
****************************************************************************************************)
METHOD m_SetMover : BOOL
VAR_INPUT
	vi_un_Index							: UINT;	// [-] 0..m_SetMoverCount - 1
	vi_udn_Id							: UDINT;	// [-] unique within the gantry, > 0
	vi_lr_Position						: LREAL;	// [mm] along the track
	vi_lr_X								: LREAL;	// [mm] X axis
	vi_b_GripperActive					: BOOL;	// used only when no fingers are configured
	(* Finger poses absolute in the MCS and grip states, index 0 = finger 1; entries beyond the finger count are ignored. *)
	vi_FingerStates						: ARRAY[0..VISU_GlobalConst_Param.VISU_un_MAX_FINGERS - 1] OF ST_VisuFingerState;
	vi_b_Fault							: BOOL := FALSE;	// TRUE: this mover is in a fault
	vi_str_FaultMessage					: STRING(80) := '';	// shown to the operator; empty shows 'Fault'
END_VAR
m_SetMover := vi_un_Index < vo_Visu.stState.nMoverCount;
IF m_SetMover THEN
	vo_Visu.stState.aMovers[vi_un_Index].nId := vi_udn_Id;
	vo_Visu.stState.aMovers[vi_un_Index].bValid := TRUE;
	vo_Visu.stState.aMovers[vi_un_Index].fPosition := vi_lr_Position;
	vo_Visu.stState.aMovers[vi_un_Index].fX := vi_lr_X;
	vo_Visu.stState.aMovers[vi_un_Index].bGripperActive := vi_b_GripperActive;
	vo_Visu.stState.aMovers[vi_un_Index].aFingerStates := vi_FingerStates;
	vo_Visu.stState.aMovers[vi_un_Index].stFault.bActive := vi_b_Fault;
	vo_Visu.stState.aMovers[vi_un_Index].stFault.sMessage := vi_str_FaultMessage;
	vo_Visu.stState.nTimestamp := m_DcTime();
END_IF
END_METHOD

